(* CODESYS project Syn_Config_2.1.0.library
   Description: Parameter sets the RPP configurator writes and the application takes over (ADR 0017).
   Version: 2.1.0.0
   Title: SynConfig
   Placeholder: SynConfig
   Company: Syntegon Group
   DefaultNamespace: SynConfig

Project tree, tasks and I/O mapping:
  libraries: SynVisu, * (Syntegon Group); Tc2_Standard, * (Beckhoff Automation GmbH)
  DUTs/
    data type E_ConfigAction
    data type E_ConfigCommand
    data type E_ConfigCommandResult
    data type E_ConfigFieldType
    data type E_ConfigResult
    data type ST_ConfigBodyComponent
    data type ST_ConfigBodyComponentParam
    data type ST_ConfigBodyComponentSet
    data type ST_ConfigCartesian
    data type ST_ConfigCartesianParam
    data type ST_ConfigCartesianSet
    data type ST_ConfigCommand
    data type ST_ConfigCommandStatus
    data type ST_ConfigConveyor
    data type ST_ConfigConveyorParam
    data type ST_ConfigConveyorSet
    data type ST_ConfigDelta
    data type ST_ConfigDeltaParam
    data type ST_ConfigDeltaSet
    data type ST_ConfigMachine
    data type ST_ConfigManifest
    data type ST_ConfigManifestEntry
    data type ST_ConfigRecipeField
    data type ST_ConfigRecipeSet
    data type ST_ConfigStaging
    data type ST_ConfigStatus
    data type ST_ConfigXtsGantry
    data type ST_ConfigXtsGantryParam
    data type ST_ConfigXtsGantrySet
    data type ST_ConfigXtsLoop
    data type ST_ConfigXtsLoopParam
    data type ST_ConfigXtsLoopSet
  GVLs/
    global variables CONFIG_GlobalConst
    global variables CONFIG_GlobalConst_Param
  POUs/
    function block _FB_ConfigBodyComponent [ST]: m_Active, m_Cycle, m_PassOnBody, m_Pose
    function block _FB_ConfigCartesian [ST]: m_Active, m_ComponentType, m_Cycle, m_Invalid, m_PassOn, m_Pose
    function block _FB_ConfigComponent [ST]: m_ComponentType, m_Handled, m_Id, m_InvalidFingers, m_InvalidModules, m_InvalidZones, m_PassOnFingers, m_PassOnLimitAreas, m_PassOnModules, m_PassOnZones, m_Register, m_Staging, m_SymbolPath
    function block _FB_ConfigConveyor [ST]: m_Active, m_ComponentType, m_Cycle, m_Invalid, m_PassOn, m_Pose
    function block _FB_ConfigDelta [ST]: m_Active, m_ComponentType, m_Cycle, m_Invalid, m_PassOn, m_Pose, m_Zone, m_ZoneCount
    function block _FB_ConfigMachine [ST]: m_AnswerCommand, m_Command, m_Cycle, m_DeclareField, m_Integer, m_Invalid, m_SetChoice, m_Switch, m_Value
    function block _FB_ConfigSensor [ST]: m_ComponentType, m_PassOn
    function block _FB_ConfigStation [ST]: m_ComponentType, m_PassOn
    function block _FB_ConfigVision [ST]: m_ComponentType, m_PassOn
    function block _FB_ConfigXtsGantry [ST]: m_Active, m_ComponentType, m_Cycle, m_Invalid, m_PassOn, m_Pose
    function block _FB_ConfigXtsLoop [ST]: m_Active, m_ComponentType, m_Cycle, m_Invalid, m_PassOn, m_Pose
    function _FC_GetVersionSynConfig [ST]
*)

// DUTs/E_ConfigAction
{attribute 'qualified_only'}
{attribute 'strict'}
TYPE E_ConfigAction :
(
	(* What a parameter FB does with its staging this cycle (internal). *)
	NONE := 0,
	TAKE_OVER := 1,	// check the staged set and take it over
	RESET := 2		// make the active set invalid: the program values apply again
) UINT;
END_TYPE

// DUTs/E_ConfigCommand
{attribute 'qualified_only'}
{attribute 'strict'}
TYPE E_ConfigCommand :
(
	(* What a machine command asks the application (config protocol 3). Values are part of the gateway contract:
	   append, never renumber. *)
	NONE := 0,
	START := 1,
	STOP := 2,
	RESET := 3
) UINT;
END_TYPE

// DUTs/E_ConfigCommandResult
{attribute 'qualified_only'}
{attribute 'strict'}
TYPE E_ConfigCommandResult :
(
	(* What the application made of the last machine command. Values are part of the gateway contract: append, never
	   renumber. *)
	NONE := 0,		// nothing asked since the PLC started
	ACCEPTED := 1,
	REJECTED := 2	// ST_ConfigCommandStatus.sMessage says why
) UINT;
END_TYPE

// DUTs/E_ConfigFieldType
{attribute 'qualified_only'}
{attribute 'strict'}
TYPE E_ConfigFieldType :
(
	(* How a recipe field's value is kept (config protocol 3). Every value travels as LREAL. Values are part of the
	   gateway contract: append, never renumber. *)
	NUMBER := 0,	// any number within fMin..fMax
	INTEGER := 1,	// a whole number within fMin..fMax, e.g. picks per cycle
	SWITCH := 2,	// on or off: 1 or 0
	CHOICE := 3		// one of the named choices: 0..nChoiceCount-1
) UINT;
END_TYPE

// DUTs/E_ConfigResult
{attribute 'qualified_only'}
{attribute 'strict'}
TYPE E_ConfigResult :
(
	(* What became of the last staged parameter set. Values are part of the gateway contract: append, never renumber. *)
	NONE := 0,		// nothing staged since the PLC started
	PENDING := 1,	// staged, waiting for the application to allow taking it over
	APPLIED := 2,	// taken over (or reset to the program values)
	REJECTED := 3	// not taken over; ST_ConfigStatus.sMessage says why
) UINT;
END_TYPE

// DUTs/ST_ConfigBodyComponent
TYPE ST_ConfigBodyComponent :
STRUCT
	(* vo_Config of _FB_ConfigVision, _FB_ConfigSensor and _FB_ConfigStation: the gateway writes stStaging and
	   stStaged, reads stStatus and stActive. *)
	stStaging : ST_ConfigStaging;
	stStaged : ST_ConfigBodyComponentParam;
	stStatus : ST_ConfigStatus;
	stActive : ST_ConfigBodyComponentParam; // effective values: the active set while one is valid, else the program values
END_STRUCT
END_TYPE

// DUTs/ST_ConfigBodyComponentParam
TYPE ST_ConfigBodyComponentParam :
STRUCT
	(* The parameter set of a component drawn from its bodies (vision system, product sensor, station): what the
	   configurator writes, never its bodies (hardware). Members as in SynVisu.ST_VisuDetectorConfig. *)
	stPose : SynVisu.ST_VisuPose; // MCS
	stOriginShift : SynVisu.ST_VisuPosition; // mm in the component's local frame
	nZoneCount : UINT;
	aZones : ARRAY[0..SynVisu.VISU_GlobalConst_Param.VISU_un_MAX_ZONES - 1] OF SynVisu.ST_VisuZone;
END_STRUCT
END_TYPE

// DUTs/ST_ConfigBodyComponentSet
TYPE ST_ConfigBodyComponentSet :
STRUCT
	(* The active parameter set of a vision system, product sensor or station as the application keeps it, in a
	   VAR PERSISTENT variable passed to m_Cycle of _FB_ConfigVision, _FB_ConfigSensor or _FB_ConfigStation. *)
	bValid : BOOL; // FALSE: no set active, the program values apply
	nVersion : UDINT; // version of stParam
	nLastVersion : UDINT; // last version handed out; versions never repeat, also after a reset
	stParam : ST_ConfigBodyComponentParam;
END_STRUCT
END_TYPE

// DUTs/ST_ConfigCartesian
TYPE ST_ConfigCartesian :
STRUCT
	(* vo_Config of _FB_ConfigCartesian: the gateway writes stStaging and stStaged, reads stStatus and stActive. *)
	stStaging : ST_ConfigStaging;
	stStaged : ST_ConfigCartesianParam;
	stStatus : ST_ConfigStatus;
	stActive : ST_ConfigCartesianParam; // effective values: the active set while one is valid, else the program values
END_STRUCT
END_TYPE

// DUTs/ST_ConfigCartesianParam
TYPE ST_ConfigCartesianParam :
STRUCT
	(* A Cartesian robot's parameter set: what the configurator writes, never its axes, strokes or rail height
	   (hardware). Members as in SynVisu.ST_VisuCartesianConfig. *)
	stPose : SynVisu.ST_VisuPose; // MCS, axis origin X = Y = 0 with Z up
	stOriginShift : SynVisu.ST_VisuPosition; // mm in the robot's local frame
	nZoneCount : UINT;
	aZones : ARRAY[0..SynVisu.VISU_GlobalConst_Param.VISU_un_MAX_ZONES - 1] OF SynVisu.ST_VisuZone;
	nFingerCount : UINT; // gripper fingers with their flange offsets (config protocol 2, ADR 0018)
	aFingers : ARRAY[0..SynVisu.VISU_GlobalConst_Param.VISU_un_MAX_FINGERS - 1] OF SynVisu.ST_VisuFinger;
	stLimitArea : SynVisu.ST_VisuLimitArea; // bActive = FALSE: none
	stTcpLimitArea : SynVisu.ST_VisuLimitArea; // bActive = FALSE: none
END_STRUCT
END_TYPE

// DUTs/ST_ConfigCartesianSet
TYPE ST_ConfigCartesianSet :
STRUCT
	(* A Cartesian robot's active parameter set as the application keeps it, in a VAR PERSISTENT variable passed to
	   _FB_ConfigCartesian.m_Cycle. *)
	bValid : BOOL; // FALSE: no set active, the program values apply
	nVersion : UDINT; // version of stParam
	nLastVersion : UDINT; // last version handed out; versions never repeat, also after a reset
	stParam : ST_ConfigCartesianParam;
END_STRUCT
END_TYPE

// DUTs/ST_ConfigCommand
TYPE ST_ConfigCommand :
STRUCT
	(* A machine command, written by the gateway with bRequested last (config protocol 3). The machine FB clears
	   bRequested once the application answered it. *)
	nCommandId : UDINT; // chosen by the gateway; ST_ConfigCommandStatus.nHandledCommandId names it once answered
	eCommand : E_ConfigCommand;
	bRequested : BOOL; // TRUE: the command waits for the application's answer
END_STRUCT
END_TYPE

// DUTs/ST_ConfigCommandStatus
TYPE ST_ConfigCommandStatus :
STRUCT
	nHandledCommandId : UDINT; // nCommandId of the last command the application answered
	eResult : E_ConfigCommandResult; // what the application made of it
	sMessage : STRING(80); // why it was rejected; empty otherwise
END_STRUCT
END_TYPE

// DUTs/ST_ConfigConveyor
TYPE ST_ConfigConveyor :
STRUCT
	(* vo_Config of _FB_ConfigConveyor: the gateway writes stStaging and stStaged, reads stStatus and stActive. *)
	stStaging : ST_ConfigStaging;
	stStaged : ST_ConfigConveyorParam;
	stStatus : ST_ConfigStatus;
	stActive : ST_ConfigConveyorParam; // effective values: the active set while one is valid, else the program values
END_STRUCT
END_TYPE

// DUTs/ST_ConfigConveyorParam
TYPE ST_ConfigConveyorParam :
STRUCT
	(* A conveyor's parameter set: what the configurator writes, never the belt's length or width (hardware).
	   Members as in SynVisu.ST_VisuConveyorConfig. *)
	stPose : SynVisu.ST_VisuPose; // MCS, belt start on the belt surface; local +X = conveying direction
	stOriginShift : SynVisu.ST_VisuPosition; // mm in the local frame from stPose: origin of the belt coordinates
	nProductTypeCount : UINT;
	aProductTypes : ARRAY[0..SynVisu.VISU_GlobalConst_Param.VISU_un_MAX_PRODUCT_TYPES - 1] OF SynVisu.ST_VisuProductType;
END_STRUCT
END_TYPE

// DUTs/ST_ConfigConveyorSet
TYPE ST_ConfigConveyorSet :
STRUCT
	(* A conveyor's active parameter set as the application keeps it, in a VAR PERSISTENT variable passed to
	   _FB_ConfigConveyor.m_Cycle. *)
	bValid : BOOL; // FALSE: no set active, the program values apply
	nVersion : UDINT; // version of stParam
	nLastVersion : UDINT; // last version handed out; versions never repeat, also after a reset
	stParam : ST_ConfigConveyorParam;
END_STRUCT
END_TYPE

// DUTs/ST_ConfigDelta
TYPE ST_ConfigDelta :
STRUCT
	(* vo_Config of _FB_ConfigDelta: the gateway writes stStaging and stStaged, reads stStatus and stActive. *)
	stStaging : ST_ConfigStaging;
	stStaged : ST_ConfigDeltaParam;
	stStatus : ST_ConfigStatus;
	stActive : ST_ConfigDeltaParam; // effective values: the active set while one is valid, else the program values
END_STRUCT
END_TYPE

// DUTs/ST_ConfigDeltaParam
TYPE ST_ConfigDeltaParam :
STRUCT
	(* A Delta robot's parameter set: what the configurator writes, never its arm geometry (hardware).
	   Members as in SynVisu.ST_VisuDeltaConfig. *)
	stPose : SynVisu.ST_VisuPose; // MCS, base centre
	stOriginShift : SynVisu.ST_VisuPosition; // mm in the base's local frame
	nZoneCount : UINT;
	aZones : ARRAY[0..SynVisu.VISU_GlobalConst_Param.VISU_un_MAX_ZONES - 1] OF SynVisu.ST_VisuZone;
	nFingerCount : UINT; // gripper fingers with their flange offsets (config protocol 2, ADR 0018)
	aFingers : ARRAY[0..SynVisu.VISU_GlobalConst_Param.VISU_un_MAX_FINGERS - 1] OF SynVisu.ST_VisuFinger;
	stWorkingArea : SynVisu.ST_VisuWorkingArea;
	stLimitArea : SynVisu.ST_VisuLimitArea; // bActive = FALSE: none
	stTcpLimitArea : SynVisu.ST_VisuLimitArea; // bActive = FALSE: none
END_STRUCT
END_TYPE

// DUTs/ST_ConfigDeltaSet
TYPE ST_ConfigDeltaSet :
STRUCT
	(* A Delta robot's active parameter set as the application keeps it, in a VAR PERSISTENT variable passed to
	   _FB_ConfigDelta.m_Cycle. *)
	bValid : BOOL; // FALSE: no set active, the program values apply
	nVersion : UDINT; // version of stParam
	nLastVersion : UDINT; // last version handed out; versions never repeat, also after a reset
	stParam : ST_ConfigDeltaParam;
END_STRUCT
END_TYPE

// DUTs/ST_ConfigMachine
TYPE ST_ConfigMachine :
STRUCT
	(* vo_Config of _FB_ConfigMachine (config protocol 3, ADR 0022), listed in the config manifest with id 0 and type
	   NONE. The gateway reads the declared fields once, writes stStaging with aStaged (bStaged or bReset last) and
	   stCommand (bRequested last), and reads stStatus, aActive and stCommandStatus every cycle. Values are kept by
	   field index, every type as LREAL (SWITCH 0 / 1, INTEGER and CHOICE whole numbers). *)
	nFieldCount : UINT; // fields [0..nFieldCount-1] are declared
	aFields : ARRAY[0..CONFIG_GlobalConst_Param.CONFIG_un_MAX_RECIPE_FIELDS - 1] OF ST_ConfigRecipeField;
	stStaging : ST_ConfigStaging;
	aStaged : ARRAY[0..CONFIG_GlobalConst_Param.CONFIG_un_MAX_RECIPE_FIELDS - 1] OF LREAL; // the proposed recipe
	stStatus : ST_ConfigStatus;
	aActive : ARRAY[0..CONFIG_GlobalConst_Param.CONFIG_un_MAX_RECIPE_FIELDS - 1] OF LREAL; // effective values
	stCommand : ST_ConfigCommand;
	stCommandStatus : ST_ConfigCommandStatus;
END_STRUCT
END_TYPE

// DUTs/ST_ConfigManifest
TYPE ST_ConfigManifest :
STRUCT
	(* Where the gateway finds the parameter FBs (ADR 0017). The application declares one instance at the symbol
	   GVL_Config.stManifest; every parameter FB registers itself with m_Register. *)
	nProtocolVersion : UINT := CONFIG_GlobalConst.CONFIG_un_PROTOCOL_VERSION;
	sLibraryVersion : STRING(15); // version of the Syn_Config library actually running, e.g. '1.0.0'
	nCount : UINT; // entries [0..nCount-1] are evaluated
	aEntries : ARRAY[0..CONFIG_GlobalConst_Param.CONFIG_un_MAX_MANIFEST_ENTRIES - 1] OF ST_ConfigManifestEntry;
END_STRUCT
END_TYPE

// DUTs/ST_ConfigManifestEntry
TYPE ST_ConfigManifestEntry :
STRUCT
	nId : UDINT; // manifest id of the Syn_Visu component the parameter FB is for
	eType : SynVisu.E_VisuComponentType; // type of that component
	sPath : STRING(255); // symbol path of the parameter FB's vo_Config, e.g. 'P_Line.fb_InfeedParam.vo_Config'
END_STRUCT
END_TYPE

// DUTs/ST_ConfigRecipeField
TYPE ST_ConfigRecipeField :
STRUCT
	(* One field of the machine's recipe as the application declares it with _FB_ConfigMachine.m_DeclareField
	   (config protocol 3, ADR 0022). The gateway reads the declarations once at discovery. *)
	sName : STRING(31); // unique in the recipe, e.g. 'BeltSpeed'
	nGroup : UDINT; // manifest id of the Syn_Visu component the field belongs to, 0 = the whole machine
	eType : E_ConfigFieldType;
	sUnit : STRING(15); // e.g. 'mm/s', '' = none
	fMin : LREAL; // smallest value of a NUMBER or INTEGER field
	fMax : LREAL; // largest value of a NUMBER or INTEGER field
	fProgramValue : LREAL; // the application's own value, which applies while no recipe is active
	nChoiceCount : UINT; // named values of a CHOICE field
	aChoices : ARRAY[0..CONFIG_GlobalConst_Param.CONFIG_un_MAX_CHOICES - 1] OF STRING(31); // their names, from value 0
END_STRUCT
END_TYPE

// DUTs/ST_ConfigRecipeSet
TYPE ST_ConfigRecipeSet :
STRUCT
	(* The machine's active recipe as the application keeps it, in a VAR PERSISTENT variable passed to
	   _FB_ConfigMachine.m_Cycle. Values by field index: keep the fields' order, add new ones at the end. *)
	bValid : BOOL; // FALSE: no recipe active, the program values apply
	nVersion : UDINT; // version of aValues
	nLastVersion : UDINT; // last version handed out; versions never repeat, also after a reset
	aValues : ARRAY[0..CONFIG_GlobalConst_Param.CONFIG_un_MAX_RECIPE_FIELDS - 1] OF LREAL;
END_STRUCT
END_TYPE

// DUTs/ST_ConfigStaging
TYPE ST_ConfigStaging :
STRUCT
	(* Written by the gateway in one ADS sum-write, bStaged or bReset last, so a set is never seen staged half
	   written (ADR 0017). The parameter FB clears bStaged and bReset once it handled them. *)
	nBaseVersion : UDINT; // active version the staged set is based on; another active version rejects it
	nStageId : UDINT; // chosen by the gateway; ST_ConfigStatus.nHandledStageId names it once handled
	bReset : BOOL; // TRUE: make the active set invalid, the program values apply again
	bStaged : BOOL; // TRUE: stStaged is complete and waits to be taken over
END_STRUCT
END_TYPE

// DUTs/ST_ConfigStatus
TYPE ST_ConfigStatus :
STRUCT
	nActiveVersion : UDINT; // version of the active set; 0 while the program values apply
	nHandledStageId : UDINT; // nStageId of the last staging handled (taken over, rejected or reset)
	eResult : E_ConfigResult; // what became of it
	sMessage : STRING(80); // why it was rejected; empty otherwise
END_STRUCT
END_TYPE

// DUTs/ST_ConfigXtsGantry
TYPE ST_ConfigXtsGantry :
STRUCT
	(* vo_Config of _FB_ConfigXtsGantry: the gateway writes stStaging and stStaged, reads stStatus and stActive. *)
	stStaging : ST_ConfigStaging;
	stStaged : ST_ConfigXtsGantryParam;
	stStatus : ST_ConfigStatus;
	stActive : ST_ConfigXtsGantryParam; // effective values: the active set while one is valid, else the program values
END_STRUCT
END_TYPE

// DUTs/ST_ConfigXtsGantryParam
TYPE ST_ConfigXtsGantryParam :
STRUCT
	(* An XTS gantry's parameter set: what the configurator writes, never its strokes, tool offsets or mover size
	   (hardware). Members as in SynVisu.ST_VisuXtsGantryConfig. *)
	stPose : SynVisu.ST_VisuPose; // MCS, track start on top of the movers with Z = 0
	stOriginShift : SynVisu.ST_VisuPosition; // mm in the track's local frame
	nModuleCount : UINT;
	aModules : ARRAY[0..SynVisu.VISU_GlobalConst_Param.VISU_un_MAX_MODULES - 1] OF SynVisu.ST_VisuTrackModule;
	nZoneCount : UINT;
	aZones : ARRAY[0..SynVisu.VISU_GlobalConst_Param.VISU_un_MAX_ZONES - 1] OF SynVisu.ST_VisuZone;
	nFingerCount : UINT; // gripper fingers of every mover, with their flange offsets (config protocol 2, ADR 0018)
	aFingers : ARRAY[0..SynVisu.VISU_GlobalConst_Param.VISU_un_MAX_FINGERS - 1] OF SynVisu.ST_VisuFinger;
	stLimitArea : SynVisu.ST_VisuLimitArea; // bActive = FALSE: none
	stTcpLimitArea : SynVisu.ST_VisuLimitArea; // bActive = FALSE: none
END_STRUCT
END_TYPE

// DUTs/ST_ConfigXtsGantrySet
TYPE ST_ConfigXtsGantrySet :
STRUCT
	(* An XTS gantry's active parameter set as the application keeps it, in a VAR PERSISTENT variable passed to
	   _FB_ConfigXtsGantry.m_Cycle. *)
	bValid : BOOL; // FALSE: no set active, the program values apply
	nVersion : UDINT; // version of stParam
	nLastVersion : UDINT; // last version handed out; versions never repeat, also after a reset
	stParam : ST_ConfigXtsGantryParam;
END_STRUCT
END_TYPE

// DUTs/ST_ConfigXtsLoop
TYPE ST_ConfigXtsLoop :
STRUCT
	(* vo_Config of _FB_ConfigXtsLoop: the gateway writes stStaging and stStaged, reads stStatus and stActive. *)
	stStaging : ST_ConfigStaging;
	stStaged : ST_ConfigXtsLoopParam;
	stStatus : ST_ConfigStatus;
	stActive : ST_ConfigXtsLoopParam; // effective values: the active set while one is valid, else the program values
END_STRUCT
END_TYPE

// DUTs/ST_ConfigXtsLoopParam
TYPE ST_ConfigXtsLoopParam :
STRUCT
	(* An XTS loop's parameter set: what the configurator writes, never its tool offset or mover size (hardware).
	   Members as in SynVisu.ST_VisuXtsLoopConfig. *)
	stPose : SynVisu.ST_VisuPose; // MCS, start of module 1
	stOriginShift : SynVisu.ST_VisuPosition; // mm in the loop's local frame
	nModuleCount : UINT;
	aModules : ARRAY[0..SynVisu.VISU_GlobalConst_Param.VISU_un_MAX_MODULES - 1] OF SynVisu.ST_VisuTrackModule;
	nZoneCount : UINT;
	aZones : ARRAY[0..SynVisu.VISU_GlobalConst_Param.VISU_un_MAX_ZONES - 1] OF SynVisu.ST_VisuZone;
	nFingerCount : UINT; // gripper fingers of every mover, with their flange offsets (config protocol 2, ADR 0018)
	aFingers : ARRAY[0..SynVisu.VISU_GlobalConst_Param.VISU_un_MAX_FINGERS - 1] OF SynVisu.ST_VisuFinger;
END_STRUCT
END_TYPE

// DUTs/ST_ConfigXtsLoopSet
TYPE ST_ConfigXtsLoopSet :
STRUCT
	(* An XTS loop's active parameter set as the application keeps it, in a VAR PERSISTENT variable passed to
	   _FB_ConfigXtsLoop.m_Cycle. *)
	bValid : BOOL; // FALSE: no set active, the program values apply
	nVersion : UDINT; // version of stParam
	nLastVersion : UDINT; // last version handed out; versions never repeat, also after a reset
	stParam : ST_ConfigXtsLoopParam;
END_STRUCT
END_TYPE

// GVLs/CONFIG_GlobalConst
(****************************************************************************************************<br>
© Syntegon Group.<br>
All rights reserved, also regarding any disposal, exploitation, reproduction, editing, distribution,<br>
as well as in the event of applications for industrial property rights.<br>
*****************************************************************************************************<br>
DESCRIPTION:<br>
Global constants of the Syn_Config library.<br>
****************************************************************************************************)
{attribute 'qualified_only'}
VAR_GLOBAL CONSTANT
	(* Version of the Syn_Config <-> gateway contract (ADR 0017). The gateway writes nothing to a PLC whose config
	   manifest reports a version it does not know (it knows 2 and 3). Bump together with CONFIG_PROTOCOL_VERSION in
	   the gateway.
	   1: conveyor (pose, origin shift, product types) and Delta (pose, origin shift, zones, working, limit and
	      TCP limit area); since library 1.1.0 also XTS gantry, XTS loop, Cartesian, vision, sensor and station
	      (new parameter FBs only: no change for a gateway or an application of 1.0.0).
	   2: gripper fingers with their flange offsets (nFingerCount, aFingers) in the parameter sets of the Delta,
	      the XTS gantry and loop and the Cartesian robot (library 2.0.0, ADR 0018).
	   3: the machine FB _FB_ConfigMachine (id 0, type NONE in the manifest): recipe fields the application declares,
	      their staging, and machine commands (library 2.1.0, ADR 0022). A PLC of version 2 still gets its parameter
	      sets written, but no recipe and no commands. *)
	CONFIG_un_PROTOCOL_VERSION			: UINT := 3;
	(* Version of this library (config manifest sLibraryVersion). Bump together with _FC_GetVersionSynConfig and the
	   project version. *)
	CONFIG_str_LIBRARY_VERSION			: STRING(15) := '2.1.0';
END_VAR

// GVLs/CONFIG_GlobalConst_Param
(****************************************************************************************************<br>
© Syntegon Group.<br>
All rights reserved, also regarding any disposal, exploitation, reproduction, editing, distribution,<br>
as well as in the event of applications for industrial property rights.<br>
*****************************************************************************************************<br>
DESCRIPTION:<br>
Library parameters of Syn_Config: array sizes of the interface structures. The lists of a parameter set have the
sizes of Syn_Visu's (VISU_GlobalConst_Param), so every set fits the visualisation it is passed on to.<br>
****************************************************************************************************)
{attribute 'qualified_only'}
VAR_GLOBAL CONSTANT
	CONFIG_un_MAX_MANIFEST_ENTRIES		: UINT := 32;	// [-] parameter FBs in the config manifest
	CONFIG_un_MAX_RECIPE_FIELDS			: UINT := 64;	// [-] fields of the machine's recipe (_FB_ConfigMachine)
	CONFIG_un_MAX_CHOICES				: UINT := 8;	// [-] named values of a CHOICE recipe field
END_VAR

// POUs/_FB_ConfigBodyComponent
(****************************************************************************************************<br>
© Syntegon Group.<br>
All rights reserved, also regarding any disposal, exploitation, reproduction, editing, distribution,<br>
as well as in the event of applications for industrial property rights.<br>
*****************************************************************************************************<br>
DESCRIPTION:<br>
Base of the parameter FBs of components drawn from their bodies (_FB_ConfigVision, _FB_ConfigSensor,<br>
_FB_ConfigStation, ADR 0017): their pose, origin shift and zones, written by the configurator, taken over when<br>
the application allows it. The bodies are hardware and stay the application's. Typical cycle:<br>
  fb_VisionParam.m_Register(vio_Manifest := GVL_Config.stManifest, vi_udn_Id := fb_Vision.m_Id());<br>
  fb_VisionParam.m_Cycle(vio_Default := VisionDefault, vio_Set := VisionSet, vi_b_ApplyAllowed := b_Stopped);<br>
  fb_Vision.m_Configure(vi_Pose := fb_VisionParam.m_Pose(), vi_lr_FieldLength := 400, ...);<br>
  fb_VisionParam.m_PassOn(vio_Visu := fb_Vision);<br>
Not used directly.<br>
*****************************************************************************************************<br>
OUTPUT VALUES:<br>
vo_Config is the contract structure the gateway reads and writes at the path in the config manifest.<br>
*****************************************************************************************************<br>
VERSION         ¦ DATE       ¦ NAME      ¦ CHANGE<br>
Syn_Config 1.1.0 ¦ 2026-11-10 ¦ J.Willner ¦ New<br>
****************************************************************************************************)
FUNCTION_BLOCK ABSTRACT _FB_ConfigBodyComponent EXTENDS _FB_ConfigComponent
VAR_OUTPUT
	vo_Config							: ST_ConfigBodyComponent;	// contract structure of the gateway
END_VAR

(****************************************************************************************************<br>
© Syntegon Group.<br>
All rights reserved, also regarding any disposal, exploitation, reproduction, editing, distribution,<br>
as well as in the event of applications for industrial property rights.<br>
*****************************************************************************************************<br>
DESCRIPTION:<br>
All effective values (zones, ...), for the application's own logic.<br>
****************************************************************************************************)
METHOD m_Active : ST_ConfigBodyComponentParam
m_Active := vo_Config.stActive;
END_METHOD

(****************************************************************************************************<br>
© Syntegon Group.<br>
All rights reserved, also regarding any disposal, exploitation, reproduction, editing, distribution,<br>
as well as in the event of applications for industrial property rights.<br>
*****************************************************************************************************<br>
DESCRIPTION:<br>
Every cycle: handles a staged set or a reset (a set only while vi_b_ApplyAllowed), keeps the active set in<br>
vio_Set and gives the effective values in vo_Config.stActive: the active set while one is valid, else the<br>
program values vio_Default.<br>
*****************************************************************************************************<br>
OUTPUT VALUES:<br>
TRUE in the cycle a set was taken over or reset.<br>
****************************************************************************************************)
METHOD m_Cycle : BOOL
VAR_IN_OUT CONSTANT
	vio_Default							: ST_ConfigBodyComponentParam;	// the application's program values
END_VAR
VAR_IN_OUT
	vio_Set								: ST_ConfigBodyComponentSet;	// the application's VAR PERSISTENT active set
END_VAR
VAR_INPUT
	vi_b_ApplyAllowed					: BOOL;	// [-] a staged set may be taken over now, e.g. while the machine stands
END_VAR
VAR
	str_TempRejection					: STRING(80);
END_VAR
m_Cycle := FALSE;
CASE m_Staging(vio_Staging := vo_Config.stStaging, vio_Status := vo_Config.stStatus, vi_b_ApplyAllowed := vi_b_ApplyAllowed,
	vi_udn_ActiveVersion := SEL(vio_Set.bValid, 0, vio_Set.nVersion)) OF
	E_ConfigAction.RESET:
		vio_Set.bValid := FALSE;
		m_Handled(vio_Staging := vo_Config.stStaging, vio_Status := vo_Config.stStatus, vi_str_Rejection := '');
		m_Cycle := TRUE;
	E_ConfigAction.TAKE_OVER:
		str_TempRejection := m_InvalidZones(vio_aZones := vo_Config.stStaged.aZones, vi_un_Count := vo_Config.stStaged.nZoneCount);
		IF str_TempRejection = '' THEN
			vio_Set.nLastVersion := vio_Set.nLastVersion + 1;
			vio_Set.nVersion := vio_Set.nLastVersion;
			vio_Set.stParam := vo_Config.stStaged;
			vio_Set.bValid := TRUE;
			m_Cycle := TRUE;
		END_IF
		m_Handled(vio_Staging := vo_Config.stStaging, vio_Status := vo_Config.stStatus, vi_str_Rejection := str_TempRejection);
END_CASE


(****************************************************************************************************
EFFECTIVE VALUES
****************************************************************************************************)
IF vio_Set.bValid THEN
	vo_Config.stActive := vio_Set.stParam;
	vo_Config.stStatus.nActiveVersion := vio_Set.nVersion;
ELSE
	vo_Config.stActive := vio_Default;
	vo_Config.stStatus.nActiveVersion := 0;
END_IF
END_METHOD

(****************************************************************************************************<br>
© Syntegon Group.<br>
All rights reserved, also regarding any disposal, exploitation, reproduction, editing, distribution,<br>
as well as in the event of applications for industrial property rights.<br>
*****************************************************************************************************<br>
DESCRIPTION:<br>
Passes the effective origin shift and zones on to the component's Syn_Visu FB; for m_PassOn of the derived FB,<br>
which knows where the visualisation keeps its zone count.<br>
****************************************************************************************************)
METHOD PROTECTED m_PassOnBody : BOOL
VAR_IN_OUT
	vio_Visu							: SynVisu._FB_VisuBodyComponent;	// the component's Syn_Visu FB
END_VAR
VAR_INPUT
	vi_un_VisuZoneCount					: UINT;	// [-] zones the visualisation has now, its stConfig.nZoneCount
END_VAR
m_PassOnBody := TRUE;
vio_Visu.m_SetOriginShift(vi_lr_X := vo_Config.stActive.stOriginShift.fX, vi_lr_Y := vo_Config.stActive.stOriginShift.fY,
	vi_lr_Z := vo_Config.stActive.stOriginShift.fZ);
m_PassOnZones(vio_Visu := vio_Visu, vio_aZones := vo_Config.stActive.aZones, vi_un_Count := vo_Config.stActive.nZoneCount,
	vi_un_VisuCount := vi_un_VisuZoneCount);
END_METHOD

(****************************************************************************************************<br>
© Syntegon Group.<br>
All rights reserved, also regarding any disposal, exploitation, reproduction, editing, distribution,<br>
as well as in the event of applications for industrial property rights.<br>
*****************************************************************************************************<br>
DESCRIPTION:<br>
Effective pose (MCS), for the application's logic and its Syn_Visu m_Configure call.<br>
****************************************************************************************************)
METHOD m_Pose : SynVisu.ST_VisuPose
m_Pose := vo_Config.stActive.stPose;
END_METHOD

END_FUNCTION_BLOCK

// POUs/_FB_ConfigVision
(****************************************************************************************************<br>
© Syntegon Group.<br>
All rights reserved, also regarding any disposal, exploitation, reproduction, editing, distribution,<br>
as well as in the event of applications for industrial property rights.<br>
*****************************************************************************************************<br>
DESCRIPTION:<br>
Parameter set of one vision system (ADR 0017): its pose, origin shift and zones. See _FB_ConfigBodyComponent.<br>
*****************************************************************************************************<br>
VERSION         ¦ DATE       ¦ NAME      ¦ CHANGE<br>
Syn_Config 1.1.0 ¦ 2026-11-10 ¦ J.Willner ¦ New<br>
****************************************************************************************************)
FUNCTION_BLOCK _FB_ConfigVision EXTENDS _FB_ConfigBodyComponent

(****************************************************************************************************<br>
© Syntegon Group.<br>
All rights reserved, also regarding any disposal, exploitation, reproduction, editing, distribution,<br>
as well as in the event of applications for industrial property rights.<br>
*****************************************************************************************************<br>
DESCRIPTION:<br>
A vision system.<br>
****************************************************************************************************)
METHOD PROTECTED m_ComponentType : SynVisu.E_VisuComponentType
m_ComponentType := SynVisu.E_VisuComponentType.VISION;
END_METHOD

(****************************************************************************************************<br>
© Syntegon Group.<br>
All rights reserved, also regarding any disposal, exploitation, reproduction, editing, distribution,<br>
as well as in the event of applications for industrial property rights.<br>
*****************************************************************************************************<br>
DESCRIPTION:<br>
Passes the effective origin shift and zones on to the vision system's Syn_Visu FB. The pose goes with the<br>
application's own m_Configure call (with the field of view, hardware): vi_Pose := m_Pose(). Call it after<br>
m_Cycle, every cycle.<br>
****************************************************************************************************)
METHOD m_PassOn : BOOL
VAR_IN_OUT
	vio_Visu							: SynVisu._FB_VisuVision;	// the vision system's Syn_Visu FB
END_VAR
m_PassOn := m_PassOnBody(vio_Visu := vio_Visu, vi_un_VisuZoneCount := vio_Visu.vo_Visu.stConfig.nZoneCount);
END_METHOD

END_FUNCTION_BLOCK

// POUs/_FB_ConfigSensor
(****************************************************************************************************<br>
© Syntegon Group.<br>
All rights reserved, also regarding any disposal, exploitation, reproduction, editing, distribution,<br>
as well as in the event of applications for industrial property rights.<br>
*****************************************************************************************************<br>
DESCRIPTION:<br>
Parameter set of one product sensor (ADR 0017): its pose, origin shift and zones. See _FB_ConfigBodyComponent.<br>
*****************************************************************************************************<br>
VERSION         ¦ DATE       ¦ NAME      ¦ CHANGE<br>
Syn_Config 1.1.0 ¦ 2026-11-10 ¦ J.Willner ¦ New<br>
****************************************************************************************************)
FUNCTION_BLOCK _FB_ConfigSensor EXTENDS _FB_ConfigBodyComponent

(****************************************************************************************************<br>
© Syntegon Group.<br>
All rights reserved, also regarding any disposal, exploitation, reproduction, editing, distribution,<br>
as well as in the event of applications for industrial property rights.<br>
*****************************************************************************************************<br>
DESCRIPTION:<br>
A product sensor.<br>
****************************************************************************************************)
METHOD PROTECTED m_ComponentType : SynVisu.E_VisuComponentType
m_ComponentType := SynVisu.E_VisuComponentType.SENSOR;
END_METHOD

(****************************************************************************************************<br>
© Syntegon Group.<br>
All rights reserved, also regarding any disposal, exploitation, reproduction, editing, distribution,<br>
as well as in the event of applications for industrial property rights.<br>
*****************************************************************************************************<br>
DESCRIPTION:<br>
Passes the effective origin shift and zones on to the sensor's Syn_Visu FB. The pose goes with the<br>
application's own m_Configure call (with the beam length, hardware): vi_Pose := m_Pose(). Call it after<br>
m_Cycle, every cycle.<br>
****************************************************************************************************)
METHOD m_PassOn : BOOL
VAR_IN_OUT
	vio_Visu							: SynVisu._FB_VisuSensor;	// the sensor's Syn_Visu FB
END_VAR
m_PassOn := m_PassOnBody(vio_Visu := vio_Visu, vi_un_VisuZoneCount := vio_Visu.vo_Visu.stConfig.nZoneCount);
END_METHOD

END_FUNCTION_BLOCK

// POUs/_FB_ConfigStation
(****************************************************************************************************<br>
© Syntegon Group.<br>
All rights reserved, also regarding any disposal, exploitation, reproduction, editing, distribution,<br>
as well as in the event of applications for industrial property rights.<br>
*****************************************************************************************************<br>
DESCRIPTION:<br>
Parameter set of one station (reject unit, labeller, ..., ADR 0017): its pose, origin shift and zones. See<br>
_FB_ConfigBodyComponent.<br>
*****************************************************************************************************<br>
VERSION         ¦ DATE       ¦ NAME      ¦ CHANGE<br>
Syn_Config 1.1.0 ¦ 2026-11-10 ¦ J.Willner ¦ New<br>
****************************************************************************************************)
FUNCTION_BLOCK _FB_ConfigStation EXTENDS _FB_ConfigBodyComponent

(****************************************************************************************************<br>
© Syntegon Group.<br>
All rights reserved, also regarding any disposal, exploitation, reproduction, editing, distribution,<br>
as well as in the event of applications for industrial property rights.<br>
*****************************************************************************************************<br>
DESCRIPTION:<br>
A station.<br>
****************************************************************************************************)
METHOD PROTECTED m_ComponentType : SynVisu.E_VisuComponentType
m_ComponentType := SynVisu.E_VisuComponentType.STATION;
END_METHOD

(****************************************************************************************************<br>
© Syntegon Group.<br>
All rights reserved, also regarding any disposal, exploitation, reproduction, editing, distribution,<br>
as well as in the event of applications for industrial property rights.<br>
*****************************************************************************************************<br>
DESCRIPTION:<br>
Passes the effective origin shift and zones on to the station's Syn_Visu FB. The pose goes with the<br>
application's own m_Configure call: vi_Pose := m_Pose(); its bodies stay the application's (hardware). Call it<br>
after m_Cycle, every cycle.<br>
****************************************************************************************************)
METHOD m_PassOn : BOOL
VAR_IN_OUT
	vio_Visu							: SynVisu._FB_VisuStation;	// the station's Syn_Visu FB
END_VAR
m_PassOn := m_PassOnBody(vio_Visu := vio_Visu, vi_un_VisuZoneCount := vio_Visu.vo_Visu.stConfig.nZoneCount);
END_METHOD

END_FUNCTION_BLOCK

// POUs/_FB_ConfigComponent
(****************************************************************************************************<br>
© Syntegon Group.<br>
All rights reserved, also regarding any disposal, exploitation, reproduction, editing, distribution,<br>
as well as in the event of applications for industrial property rights.<br>
*****************************************************************************************************<br>
DESCRIPTION:<br>
Base of every parameter FB (_FB_ConfigConveyor, _FB_ConfigDelta, _FB_ConfigXtsGantry, ...): the config<br>
manifest entry, what is done with a staging (ADR 0017) and the helpers for zones, fingers, limit areas and<br>
track modules the derived FBs share. Not used directly.<br>
*****************************************************************************************************<br>
VERSION         ¦ DATE       ¦ NAME      ¦ CHANGE<br>
Syn_Config 1.0.0 ¦ 2026-11-10 ¦ J.Willner ¦ First version: conveyor and Delta<br>
Syn_Config 1.1.0 ¦ 2026-11-10 ¦ J.Willner ¦ Helpers m_PassOn..., m_Invalid... for every type<br>
Syn_Config 2.0.0 ¦ 2026-11-11 ¦ J.Willner ¦ m_InvalidFingers, m_PassOnFingers (ADR 0018)<br>
****************************************************************************************************)
{attribute 'reflection'}
FUNCTION_BLOCK ABSTRACT _FB_ConfigComponent
VAR
	udn_ComponentId						: UDINT;	// [-] id of the Syn_Visu component, 0 = not registered
	(* Device tree path of this instance, e.g. 'RPP_Visu.Syn_Visu_Demo.P_VisuDemoDelta.fb_InfeedParam', set by TwinCAT
	   at initialisation. *)
	{attribute 'instance-path'}
	{attribute 'noinit'}
	str_InstancePath					: STRING(255);
	str_SymbolPath						: STRING(255);	// symbol path of vo_Config for the manifest, from str_InstancePath
END_VAR

(****************************************************************************************************<br>
© Syntegon Group.<br>
All rights reserved, also regarding any disposal, exploitation, reproduction, editing, distribution,<br>
as well as in the event of applications for industrial property rights.<br>
*****************************************************************************************************<br>
DESCRIPTION:<br>
Type of the Syn_Visu component this FB parametrises. Overridden by every derived FB.<br>
****************************************************************************************************)
METHOD PROTECTED m_ComponentType : SynVisu.E_VisuComponentType
m_ComponentType := SynVisu.E_VisuComponentType.NONE;
END_METHOD

(****************************************************************************************************<br>
© Syntegon Group.<br>
All rights reserved, also regarding any disposal, exploitation, reproduction, editing, distribution,<br>
as well as in the event of applications for industrial property rights.<br>
*****************************************************************************************************<br>
DESCRIPTION:<br>
Reports the staging as handled: taken over (or reset) with an empty vi_str_Rejection, else rejected for that<br>
reason. Clears bStaged and bReset. TRUE when taken over.<br>
****************************************************************************************************)
METHOD PROTECTED m_Handled : BOOL
VAR_IN_OUT
	vio_Staging							: ST_ConfigStaging;	// vo_Config.stStaging
	vio_Status							: ST_ConfigStatus;	// vo_Config.stStatus
END_VAR
VAR_INPUT
	vi_str_Rejection					: STRING(80);	// why the set is not taken over; '' = taken over
END_VAR
m_Handled := vi_str_Rejection = '';
vio_Status.nHandledStageId := vio_Staging.nStageId;
IF m_Handled THEN
	vio_Status.eResult := E_ConfigResult.APPLIED;
	vio_Status.sMessage := '';
ELSE
	vio_Status.eResult := E_ConfigResult.REJECTED;
	vio_Status.sMessage := vi_str_Rejection;
END_IF
vio_Staging.bStaged := FALSE;
vio_Staging.bReset := FALSE;
END_METHOD

(****************************************************************************************************<br>
© Syntegon Group.<br>
All rights reserved, also regarding any disposal, exploitation, reproduction, editing, distribution,<br>
as well as in the event of applications for industrial property rights.<br>
*****************************************************************************************************<br>
DESCRIPTION:<br>
Id given to m_Register (the Syn_Visu component's id); 0 while not registered.<br>
****************************************************************************************************)
METHOD m_Id : UDINT
m_Id := udn_ComponentId;
END_METHOD

(****************************************************************************************************<br>
© Syntegon Group.<br>
All rights reserved, also regarding any disposal, exploitation, reproduction, editing, distribution,<br>
as well as in the event of applications for industrial property rights.<br>
*****************************************************************************************************<br>
DESCRIPTION:<br>
Why a staged set's gripper fingers cannot be taken over; '' when they can: more fingers than the list holds, or<br>
a finger without a diameter or height.<br>
****************************************************************************************************)
METHOD PROTECTED m_InvalidFingers : STRING(80)
VAR_IN_OUT CONSTANT
	(* staged fingers *)
	vio_aFingers						: ARRAY[0..SynVisu.VISU_GlobalConst_Param.VISU_un_MAX_FINGERS - 1] OF SynVisu.ST_VisuFinger;
END_VAR
VAR_INPUT
	vi_un_Count							: UINT;	// [-] staged fingers in vio_aFingers
END_VAR
VAR
	un_TempIndex						: UINT;
END_VAR
m_InvalidFingers := '';
IF vi_un_Count > SynVisu.VISU_GlobalConst_Param.VISU_un_MAX_FINGERS THEN
	m_InvalidFingers := CONCAT('More than ', CONCAT(UINT_TO_STRING(SynVisu.VISU_GlobalConst_Param.VISU_un_MAX_FINGERS), ' fingers'));
	RETURN;
END_IF
un_TempIndex := 0;
WHILE un_TempIndex < vi_un_Count DO
	IF vio_aFingers[un_TempIndex].fDiameter <= 0 OR vio_aFingers[un_TempIndex].fHeight <= 0 THEN
		m_InvalidFingers := CONCAT('Finger ', CONCAT(UINT_TO_STRING(un_TempIndex + 1), ' has no diameter or height'));
		RETURN;
	END_IF
	un_TempIndex := un_TempIndex + 1;
END_WHILE
END_METHOD

(****************************************************************************************************<br>
© Syntegon Group.<br>
All rights reserved, also regarding any disposal, exploitation, reproduction, editing, distribution,<br>
as well as in the event of applications for industrial property rights.<br>
*****************************************************************************************************<br>
DESCRIPTION:<br>
Why a staged set's track modules cannot be taken over; '' when they can: more modules than the list holds,<br>
none at all, or a module without a length.<br>
****************************************************************************************************)
METHOD PROTECTED m_InvalidModules : STRING(80)
VAR_IN_OUT CONSTANT
	(* staged modules *)
	vio_aModules						: ARRAY[0..SynVisu.VISU_GlobalConst_Param.VISU_un_MAX_MODULES - 1] OF SynVisu.ST_VisuTrackModule;
END_VAR
VAR_INPUT
	vi_un_Count							: UINT;	// [-] staged modules in vio_aModules
END_VAR
VAR
	un_TempIndex						: UINT;
END_VAR
m_InvalidModules := '';
IF vi_un_Count > SynVisu.VISU_GlobalConst_Param.VISU_un_MAX_MODULES THEN
	m_InvalidModules := CONCAT('More than ', CONCAT(UINT_TO_STRING(SynVisu.VISU_GlobalConst_Param.VISU_un_MAX_MODULES), ' track modules'));
	RETURN;
END_IF
IF vi_un_Count = 0 THEN
	m_InvalidModules := 'A track without modules';
	RETURN;
END_IF
un_TempIndex := 0;
WHILE un_TempIndex < vi_un_Count DO
	IF vio_aModules[un_TempIndex].fLength <= 0 THEN
		m_InvalidModules := CONCAT('Track module ', CONCAT(UINT_TO_STRING(un_TempIndex + 1), ' has no length'));
		RETURN;
	END_IF
	un_TempIndex := un_TempIndex + 1;
END_WHILE
END_METHOD

(****************************************************************************************************<br>
© Syntegon Group.<br>
All rights reserved, also regarding any disposal, exploitation, reproduction, editing, distribution,<br>
as well as in the event of applications for industrial property rights.<br>
*****************************************************************************************************<br>
DESCRIPTION:<br>
Why a staged set's zones cannot be taken over; '' when they can: more zones than the list holds, or a zone on<br>
no conveyor (id 0).<br>
****************************************************************************************************)
METHOD PROTECTED m_InvalidZones : STRING(80)
VAR_IN_OUT CONSTANT
	(* staged zones *)
	vio_aZones							: ARRAY[0..SynVisu.VISU_GlobalConst_Param.VISU_un_MAX_ZONES - 1] OF SynVisu.ST_VisuZone;
END_VAR
VAR_INPUT
	vi_un_Count							: UINT;	// [-] staged zones in vio_aZones
END_VAR
VAR
	un_TempIndex						: UINT;
END_VAR
m_InvalidZones := '';
IF vi_un_Count > SynVisu.VISU_GlobalConst_Param.VISU_un_MAX_ZONES THEN
	m_InvalidZones := CONCAT('More than ', CONCAT(UINT_TO_STRING(SynVisu.VISU_GlobalConst_Param.VISU_un_MAX_ZONES), ' zones'));
	RETURN;
END_IF
un_TempIndex := 0;
WHILE un_TempIndex < vi_un_Count DO
	IF vio_aZones[un_TempIndex].nConveyorId = 0 THEN
		m_InvalidZones := CONCAT('Zone ', CONCAT(UINT_TO_STRING(un_TempIndex + 1), ' lies on no conveyor'));
		RETURN;
	END_IF
	un_TempIndex := un_TempIndex + 1;
END_WHILE
END_METHOD

(****************************************************************************************************<br>
© Syntegon Group.<br>
All rights reserved, also regarding any disposal, exploitation, reproduction, editing, distribution,<br>
as well as in the event of applications for industrial property rights.<br>
*****************************************************************************************************<br>
DESCRIPTION:<br>
Passes the effective gripper fingers with their flange offsets on to a robot's Syn_Visu FB (ADR 0018). Syn_Visu's<br>
finger count only grows: the fingers are cleared first only when the set has fewer than the visualisation, so<br>
its config version only changes when a value does.<br>
****************************************************************************************************)
METHOD PROTECTED m_PassOnFingers : BOOL
VAR_IN_OUT
	vio_Visu							: SynVisu._FB_VisuRobot;	// the robot's Syn_Visu FB
END_VAR
VAR_IN_OUT CONSTANT
	(* effective fingers *)
	vio_aFingers						: ARRAY[0..SynVisu.VISU_GlobalConst_Param.VISU_un_MAX_FINGERS - 1] OF SynVisu.ST_VisuFinger;
END_VAR
VAR_INPUT
	vi_un_Count							: UINT;	// [-] effective fingers in vio_aFingers
	vi_un_VisuCount						: UINT;	// [-] fingers the visualisation has now, its stConfig.nFingerCount
END_VAR
VAR
	un_TempIndex						: UINT;
END_VAR
m_PassOnFingers := TRUE;
IF vi_un_VisuCount > vi_un_Count THEN
	vio_Visu.m_ClearFingers();
END_IF
un_TempIndex := 0;
WHILE un_TempIndex < vi_un_Count AND un_TempIndex < SynVisu.VISU_GlobalConst_Param.VISU_un_MAX_FINGERS DO
	vio_Visu.m_SetFinger(vi_un_Finger := un_TempIndex + 1, vi_lr_Diameter := vio_aFingers[un_TempIndex].fDiameter,
		vi_lr_Height := vio_aFingers[un_TempIndex].fHeight);
	vio_Visu.m_SetFingerOffset(vi_un_Finger := un_TempIndex + 1, vi_lr_X := vio_aFingers[un_TempIndex].stOffset.fX,
		vi_lr_Y := vio_aFingers[un_TempIndex].stOffset.fY, vi_lr_Z := vio_aFingers[un_TempIndex].stOffset.fZ,
		vi_lr_Rz := vio_aFingers[un_TempIndex].stOffset.fRz);
	un_TempIndex := un_TempIndex + 1;
END_WHILE
END_METHOD

(****************************************************************************************************<br>
© Syntegon Group.<br>
All rights reserved, also regarding any disposal, exploitation, reproduction, editing, distribution,<br>
as well as in the event of applications for industrial property rights.<br>
*****************************************************************************************************<br>
DESCRIPTION:<br>
Passes the effective limit area and TCP limit area on to a robot's Syn_Visu FB (Delta, XTS gantry, Cartesian);<br>
an area with bActive = FALSE is cleared.<br>
****************************************************************************************************)
METHOD PROTECTED m_PassOnLimitAreas : BOOL
VAR_IN_OUT
	vio_Visu							: SynVisu._FB_VisuRobot;	// the robot's Syn_Visu FB
END_VAR
VAR_IN_OUT CONSTANT
	vio_LimitArea						: SynVisu.ST_VisuLimitArea;	// effective limit area
	vio_TcpLimitArea					: SynVisu.ST_VisuLimitArea;	// effective TCP limit area
END_VAR
m_PassOnLimitAreas := TRUE;
IF vio_LimitArea.bActive THEN
	vio_Visu.m_SetLimitArea(vi_lr_XMin := vio_LimitArea.fXMin, vi_lr_XMax := vio_LimitArea.fXMax,
		vi_lr_YMin := vio_LimitArea.fYMin, vi_lr_YMax := vio_LimitArea.fYMax,
		vi_lr_ZMin := vio_LimitArea.fZMin, vi_lr_ZMax := vio_LimitArea.fZMax);
ELSE
	vio_Visu.m_ClearLimitArea();
END_IF
IF vio_TcpLimitArea.bActive THEN
	vio_Visu.m_SetTcpLimitArea(vi_lr_XMin := vio_TcpLimitArea.fXMin, vi_lr_XMax := vio_TcpLimitArea.fXMax,
		vi_lr_YMin := vio_TcpLimitArea.fYMin, vi_lr_YMax := vio_TcpLimitArea.fYMax,
		vi_lr_ZMin := vio_TcpLimitArea.fZMin, vi_lr_ZMax := vio_TcpLimitArea.fZMax);
ELSE
	vio_Visu.m_ClearTcpLimitArea();
END_IF
END_METHOD

(****************************************************************************************************<br>
© Syntegon Group.<br>
All rights reserved, also regarding any disposal, exploitation, reproduction, editing, distribution,<br>
as well as in the event of applications for industrial property rights.<br>
*****************************************************************************************************<br>
DESCRIPTION:<br>
Passes the effective track modules on to an XTS track's Syn_Visu FB (XTS gantry, XTS loop). Syn_Visu's module<br>
count only grows: the modules are cleared first only when the set has fewer than the visualisation, so its<br>
config version only changes when a value does.<br>
****************************************************************************************************)
METHOD PROTECTED m_PassOnModules : BOOL
VAR_IN_OUT
	vio_Visu							: SynVisu._FB_VisuXtsTrack;	// the track's Syn_Visu FB
END_VAR
VAR_IN_OUT CONSTANT
	(* effective modules *)
	vio_aModules						: ARRAY[0..SynVisu.VISU_GlobalConst_Param.VISU_un_MAX_MODULES - 1] OF SynVisu.ST_VisuTrackModule;
END_VAR
VAR_INPUT
	vi_un_Count							: UINT;	// [-] effective modules in vio_aModules
	vi_un_VisuCount						: UINT;	// [-] modules the visualisation has now, its stConfig.nModuleCount
END_VAR
VAR
	un_TempIndex						: UINT;
END_VAR
m_PassOnModules := TRUE;
IF vi_un_VisuCount > vi_un_Count THEN
	vio_Visu.m_ClearModules();
END_IF
un_TempIndex := 0;
WHILE un_TempIndex < vi_un_Count AND un_TempIndex < SynVisu.VISU_GlobalConst_Param.VISU_un_MAX_MODULES DO
	vio_Visu.m_SetModule(vi_un_Module := un_TempIndex + 1, vi_e_Kind := vio_aModules[un_TempIndex].eKind,
		vi_lr_Length := vio_aModules[un_TempIndex].fLength);
	un_TempIndex := un_TempIndex + 1;
END_WHILE
END_METHOD

(****************************************************************************************************<br>
© Syntegon Group.<br>
All rights reserved, also regarding any disposal, exploitation, reproduction, editing, distribution,<br>
as well as in the event of applications for industrial property rights.<br>
*****************************************************************************************************<br>
DESCRIPTION:<br>
Passes the effective zones on to a Syn_Visu component with zones (robot, detector, station). Syn_Visu's zone<br>
count only grows: the zones are cleared first only when the set has fewer than the visualisation, so its<br>
config version only changes when a value does.<br>
****************************************************************************************************)
METHOD PROTECTED m_PassOnZones : BOOL
VAR_IN_OUT
	vio_Visu							: SynVisu._FB_VisuZoneComponent;	// the component's Syn_Visu FB
END_VAR
VAR_IN_OUT CONSTANT
	(* effective zones *)
	vio_aZones							: ARRAY[0..SynVisu.VISU_GlobalConst_Param.VISU_un_MAX_ZONES - 1] OF SynVisu.ST_VisuZone;
END_VAR
VAR_INPUT
	vi_un_Count							: UINT;	// [-] effective zones in vio_aZones
	vi_un_VisuCount						: UINT;	// [-] zones the visualisation has now, its stConfig.nZoneCount
END_VAR
VAR
	un_TempIndex						: UINT;
END_VAR
m_PassOnZones := TRUE;
IF vi_un_VisuCount > vi_un_Count THEN
	vio_Visu.m_ClearZones();
END_IF
un_TempIndex := 0;
WHILE un_TempIndex < vi_un_Count AND un_TempIndex < SynVisu.VISU_GlobalConst_Param.VISU_un_MAX_ZONES DO
	vio_Visu.m_SetZone(vi_un_Zone := un_TempIndex + 1, vi_udn_ConveyorId := vio_aZones[un_TempIndex].nConveyorId,
		vi_lr_Start := vio_aZones[un_TempIndex].fStart, vi_lr_End := vio_aZones[un_TempIndex].fEnd,
		vi_lr_AllocationOffset := vio_aZones[un_TempIndex].fAllocationOffset,
		vi_lr_CcsOffset := vio_aZones[un_TempIndex].fCcsOffset,
		vi_lr_StartY := vio_aZones[un_TempIndex].fStartY, vi_lr_EndY := vio_aZones[un_TempIndex].fEndY);
	un_TempIndex := un_TempIndex + 1;
END_WHILE
END_METHOD

(****************************************************************************************************<br>
© Syntegon Group.<br>
All rights reserved, also regarding any disposal, exploitation, reproduction, editing, distribution,<br>
as well as in the event of applications for industrial property rights.<br>
*****************************************************************************************************<br>
DESCRIPTION:<br>
Adds this parameter FB to the config manifest under the id of the Syn_Visu component it parametrises.<br>
Idempotent: call it every cycle. The symbol path the gateway reads comes from the instance's own path, as in<br>
Syn_Visu (VISU_un_INSTANCE_PATH_SKIP).<br>
*****************************************************************************************************<br>
OUTPUT VALUES:<br>
FALSE for vi_udn_Id = 0 (but for _FB_ConfigMachine, which registers with id 0), an id already used by a<br>
different entry, or a full manifest.<br>
****************************************************************************************************)
METHOD m_Register : BOOL
VAR_IN_OUT
	vio_Manifest						: ST_ConfigManifest;	// GVL_Config.stManifest of the application
END_VAR
VAR_INPUT
	vi_udn_Id							: UDINT;	// [-] id of the Syn_Visu component, e.g. fb_Infeed.m_Id()
END_VAR
VAR
	e_TempType							: SynVisu.E_VisuComponentType;
	un_TempIndex						: UINT;
END_VAR
m_Register := FALSE;
(* Always report the contract version of the library actually running, also after an online change. *)
vio_Manifest.nProtocolVersion := CONFIG_GlobalConst.CONFIG_un_PROTOCOL_VERSION;
vio_Manifest.sLibraryVersion := CONFIG_GlobalConst.CONFIG_str_LIBRARY_VERSION;
e_TempType := m_ComponentType();
(* Id 0 is the machine FB's, whose type is NONE (_FB_ConfigMachine); every parameter FB has a component's id. *)
IF (vi_udn_Id = 0) <> (e_TempType = SynVisu.E_VisuComponentType.NONE) THEN
	RETURN;
END_IF
IF str_SymbolPath = '' THEN
	str_SymbolPath := m_SymbolPath();
END_IF

(* An existing entry with the same id must match exactly. *)
un_TempIndex := 0;
WHILE un_TempIndex < vio_Manifest.nCount AND un_TempIndex < CONFIG_GlobalConst_Param.CONFIG_un_MAX_MANIFEST_ENTRIES DO
	IF vio_Manifest.aEntries[un_TempIndex].nId = vi_udn_Id THEN
		m_Register := vio_Manifest.aEntries[un_TempIndex].eType = e_TempType
					AND vio_Manifest.aEntries[un_TempIndex].sPath = str_SymbolPath;
		IF m_Register THEN
			udn_ComponentId := vi_udn_Id;
		END_IF
		RETURN;
	END_IF
	un_TempIndex := un_TempIndex + 1;
END_WHILE

(* New entry. *)
IF vio_Manifest.nCount >= CONFIG_GlobalConst_Param.CONFIG_un_MAX_MANIFEST_ENTRIES THEN
	RETURN;
END_IF
vio_Manifest.aEntries[vio_Manifest.nCount].nId := vi_udn_Id;
vio_Manifest.aEntries[vio_Manifest.nCount].eType := e_TempType;
vio_Manifest.aEntries[vio_Manifest.nCount].sPath := str_SymbolPath;
vio_Manifest.nCount := vio_Manifest.nCount + 1;
udn_ComponentId := vi_udn_Id;
m_Register := TRUE;
END_METHOD

(****************************************************************************************************<br>
© Syntegon Group.<br>
All rights reserved, also regarding any disposal, exploitation, reproduction, editing, distribution,<br>
as well as in the event of applications for industrial property rights.<br>
*****************************************************************************************************<br>
DESCRIPTION:<br>
What to do with the staging this cycle: a reset at once; a staged set only while the application allows it<br>
(else the status says PENDING) and only on the active version it is based on (else it is rejected here).<br>
****************************************************************************************************)
METHOD PROTECTED m_Staging : E_ConfigAction
VAR_IN_OUT
	vio_Staging							: ST_ConfigStaging;	// vo_Config.stStaging
	vio_Status							: ST_ConfigStatus;	// vo_Config.stStatus
END_VAR
VAR_INPUT
	vi_b_ApplyAllowed					: BOOL;	// [-] the application allows taking a set over now
	vi_udn_ActiveVersion				: UDINT;	// [-] version of the active set, 0 = program values
END_VAR
m_Staging := E_ConfigAction.NONE;
IF vio_Staging.bReset THEN
	m_Staging := E_ConfigAction.RESET;
ELSIF vio_Staging.bStaged THEN
	IF NOT vi_b_ApplyAllowed THEN
		vio_Status.eResult := E_ConfigResult.PENDING;
	ELSIF vio_Staging.nBaseVersion <> vi_udn_ActiveVersion THEN
		m_Handled(vio_Staging := vio_Staging, vio_Status := vio_Status,
			vi_str_Rejection := CONCAT(CONCAT('Based on version ', UDINT_TO_STRING(vio_Staging.nBaseVersion)),
				CONCAT(', but version ', CONCAT(UDINT_TO_STRING(vi_udn_ActiveVersion), ' is active'))));
	ELSE
		m_Staging := E_ConfigAction.TAKE_OVER;
	END_IF
END_IF
END_METHOD

(****************************************************************************************************<br>
© Syntegon Group.<br>
All rights reserved, also regarding any disposal, exploitation, reproduction, editing, distribution,<br>
as well as in the event of applications for industrial property rights.<br>
*****************************************************************************************************<br>
DESCRIPTION:<br>
Symbol path of this instance's vo_Config as the gateway reads it, from the instance path TwinCAT sets: the<br>
first VISU_un_INSTANCE_PATH_SKIP segments (TwinCAT project, PLC project) are left out, '.vo_Config' is appended.<br>
E.g. 'RPP_Visu.Syn_Visu_Demo.P_VisuDemoDelta.fb_InfeedParam' -> 'P_VisuDemoDelta.fb_InfeedParam.vo_Config'.<br>
****************************************************************************************************)
METHOD PRIVATE m_SymbolPath : STRING(255)
VAR
	un_TempRead							: UINT;	// [-] byte index in str_InstancePath
	un_TempWrite						: UINT;	// [-] byte index in the result
	un_TempDots							: UINT;	// [-] dots passed
END_VAR
VAR CONSTANT
	un_MAX_INDEX						: UINT := 255;	// [-] last byte of a STRING(255), its terminating zero
	by_DOT								: BYTE := 16#2E;	// '.'
	str_SUFFIX							: STRING(15) := '.vo_Config';	// every parameter FB's contract structure
END_VAR
(* Skip the leading segments, up to and including the VISU_un_INSTANCE_PATH_SKIP-th dot. *)
un_TempRead := 0;
un_TempDots := 0;
WHILE un_TempDots < SynVisu.VISU_GlobalConst_Param.VISU_un_INSTANCE_PATH_SKIP AND un_TempRead < un_MAX_INDEX
	AND str_InstancePath[un_TempRead] <> 0
DO
	IF str_InstancePath[un_TempRead] = by_DOT THEN
		un_TempDots := un_TempDots + 1;
	END_IF
	un_TempRead := un_TempRead + 1;
END_WHILE
IF un_TempDots < SynVisu.VISU_GlobalConst_Param.VISU_un_INSTANCE_PATH_SKIP THEN
	un_TempRead := 0;
END_IF

(* The rest of the instance path, then the contract structure. *)
un_TempWrite := 0;
WHILE un_TempRead < un_MAX_INDEX AND str_InstancePath[un_TempRead] <> 0 AND un_TempWrite < un_MAX_INDEX DO
	m_SymbolPath[un_TempWrite] := str_InstancePath[un_TempRead];
	un_TempRead := un_TempRead + 1;
	un_TempWrite := un_TempWrite + 1;
END_WHILE
un_TempRead := 0;
WHILE str_SUFFIX[un_TempRead] <> 0 AND un_TempWrite < un_MAX_INDEX DO
	m_SymbolPath[un_TempWrite] := str_SUFFIX[un_TempRead];
	un_TempRead := un_TempRead + 1;
	un_TempWrite := un_TempWrite + 1;
END_WHILE
m_SymbolPath[un_TempWrite] := 0;
END_METHOD

END_FUNCTION_BLOCK

// POUs/_FB_ConfigConveyor
(****************************************************************************************************<br>
© Syntegon Group.<br>
All rights reserved, also regarding any disposal, exploitation, reproduction, editing, distribution,<br>
as well as in the event of applications for industrial property rights.<br>
*****************************************************************************************************<br>
DESCRIPTION:<br>
Parameter set of one conveyor (ADR 0017): its pose, origin shift and product types, written by the configurator,<br>
taken over when the application allows it. Typical cycle, before the Syn_Visu calls of the conveyor:<br>
  fb_InfeedParam.m_Register(vio_Manifest := GVL_Config.stManifest, vi_udn_Id := fb_Infeed.m_Id());<br>
  fb_InfeedParam.m_Cycle(vio_Default := InfeedDefault, vio_Set := InfeedSet, vi_b_ApplyAllowed := b_Stopped);<br>
  fb_Infeed.m_Configure(vi_Pose := fb_InfeedParam.m_Pose(), vi_lr_Length := 3000, vi_lr_Width := 400);<br>
  fb_InfeedParam.m_PassOn(vio_Visu := fb_Infeed);<br>
InfeedSet is the application's VAR PERSISTENT ST_ConfigConveyorSet; InfeedDefault its program values.<br>
*****************************************************************************************************<br>
OUTPUT VALUES:<br>
vo_Config is the contract structure the gateway reads and writes at the path in the config manifest.<br>
*****************************************************************************************************<br>
VERSION         ¦ DATE       ¦ NAME      ¦ CHANGE<br>
Syn_Config 1.0.0 ¦ 2026-11-10 ¦ J.Willner ¦ First version<br>
****************************************************************************************************)
FUNCTION_BLOCK _FB_ConfigConveyor EXTENDS _FB_ConfigComponent
VAR_OUTPUT
	vo_Config							: ST_ConfigConveyor;	// contract structure of the gateway
END_VAR

(****************************************************************************************************<br>
© Syntegon Group.<br>
All rights reserved, also regarding any disposal, exploitation, reproduction, editing, distribution,<br>
as well as in the event of applications for industrial property rights.<br>
*****************************************************************************************************<br>
DESCRIPTION:<br>
All effective values (origin shift, product types, ...), for the application's own logic.<br>
****************************************************************************************************)
METHOD m_Active : ST_ConfigConveyorParam
m_Active := vo_Config.stActive;
END_METHOD

(****************************************************************************************************<br>
© Syntegon Group.<br>
All rights reserved, also regarding any disposal, exploitation, reproduction, editing, distribution,<br>
as well as in the event of applications for industrial property rights.<br>
*****************************************************************************************************<br>
DESCRIPTION:<br>
A conveyor.<br>
****************************************************************************************************)
METHOD PROTECTED m_ComponentType : SynVisu.E_VisuComponentType
m_ComponentType := SynVisu.E_VisuComponentType.CONVEYOR;
END_METHOD

(****************************************************************************************************<br>
© Syntegon Group.<br>
All rights reserved, also regarding any disposal, exploitation, reproduction, editing, distribution,<br>
as well as in the event of applications for industrial property rights.<br>
*****************************************************************************************************<br>
DESCRIPTION:<br>
Every cycle: handles a staged set or a reset (a set only while vi_b_ApplyAllowed), keeps the active set in<br>
vio_Set and gives the effective values in vo_Config.stActive: the active set while one is valid, else the<br>
program values vio_Default.<br>
*****************************************************************************************************<br>
OUTPUT VALUES:<br>
TRUE in the cycle a set was taken over or reset.<br>
****************************************************************************************************)
METHOD m_Cycle : BOOL
VAR_IN_OUT CONSTANT
	vio_Default							: ST_ConfigConveyorParam;	// the application's program values
END_VAR
VAR_IN_OUT
	vio_Set								: ST_ConfigConveyorSet;	// the application's VAR PERSISTENT active set
END_VAR
VAR_INPUT
	vi_b_ApplyAllowed					: BOOL;	// [-] a staged set may be taken over now, e.g. while the machine stands
END_VAR
VAR
	str_TempRejection					: STRING(80);
END_VAR
m_Cycle := FALSE;
CASE m_Staging(vio_Staging := vo_Config.stStaging, vio_Status := vo_Config.stStatus, vi_b_ApplyAllowed := vi_b_ApplyAllowed,
	vi_udn_ActiveVersion := SEL(vio_Set.bValid, 0, vio_Set.nVersion)) OF
	E_ConfigAction.RESET:
		vio_Set.bValid := FALSE;
		m_Handled(vio_Staging := vo_Config.stStaging, vio_Status := vo_Config.stStatus, vi_str_Rejection := '');
		m_Cycle := TRUE;
	E_ConfigAction.TAKE_OVER:
		str_TempRejection := m_Invalid(vio_Param := vo_Config.stStaged);
		IF str_TempRejection = '' THEN
			vio_Set.nLastVersion := vio_Set.nLastVersion + 1;
			vio_Set.nVersion := vio_Set.nLastVersion;
			vio_Set.stParam := vo_Config.stStaged;
			vio_Set.bValid := TRUE;
			m_Cycle := TRUE;
		END_IF
		m_Handled(vio_Staging := vo_Config.stStaging, vio_Status := vo_Config.stStatus, vi_str_Rejection := str_TempRejection);
END_CASE


(****************************************************************************************************
EFFECTIVE VALUES
****************************************************************************************************)
IF vio_Set.bValid THEN
	vo_Config.stActive := vio_Set.stParam;
	vo_Config.stStatus.nActiveVersion := vio_Set.nVersion;
ELSE
	vo_Config.stActive := vio_Default;
	vo_Config.stStatus.nActiveVersion := 0;
END_IF
END_METHOD

(****************************************************************************************************<br>
© Syntegon Group.<br>
All rights reserved, also regarding any disposal, exploitation, reproduction, editing, distribution,<br>
as well as in the event of applications for industrial property rights.<br>
*****************************************************************************************************<br>
DESCRIPTION:<br>
Why a staged set cannot be taken over; '' when it can: more product types than the list holds, a product type<br>
without a number or a number used twice.<br>
****************************************************************************************************)
METHOD PRIVATE m_Invalid : STRING(80)
VAR_IN_OUT CONSTANT
	vio_Param							: ST_ConfigConveyorParam;	// the staged set
END_VAR
VAR
	un_TempIndex						: UINT;
	un_TempOther						: UINT;
END_VAR
m_Invalid := '';
IF vio_Param.nProductTypeCount > SynVisu.VISU_GlobalConst_Param.VISU_un_MAX_PRODUCT_TYPES THEN
	m_Invalid := CONCAT('More than ', CONCAT(UINT_TO_STRING(SynVisu.VISU_GlobalConst_Param.VISU_un_MAX_PRODUCT_TYPES), ' product types'));
	RETURN;
END_IF
un_TempIndex := 0;
WHILE un_TempIndex < vio_Param.nProductTypeCount DO
	IF vio_Param.aProductTypes[un_TempIndex].nId = 0 THEN
		m_Invalid := 'A product type without a number';
		RETURN;
	END_IF
	un_TempOther := 0;
	WHILE un_TempOther < un_TempIndex DO
		IF vio_Param.aProductTypes[un_TempOther].nId = vio_Param.aProductTypes[un_TempIndex].nId THEN
			m_Invalid := CONCAT('Product type ', CONCAT(UDINT_TO_STRING(vio_Param.aProductTypes[un_TempIndex].nId), ' is defined twice'));
			RETURN;
		END_IF
		un_TempOther := un_TempOther + 1;
	END_WHILE
	un_TempIndex := un_TempIndex + 1;
END_WHILE
END_METHOD

(****************************************************************************************************<br>
© Syntegon Group.<br>
All rights reserved, also regarding any disposal, exploitation, reproduction, editing, distribution,<br>
as well as in the event of applications for industrial property rights.<br>
*****************************************************************************************************<br>
DESCRIPTION:<br>
Passes the effective origin shift and product types on to the conveyor's Syn_Visu FB, so the visualisation shows<br>
what the machine uses. The pose goes with the application's own m_Configure call (with the belt's length and<br>
width, hardware): vi_Pose := m_Pose(). Call it after m_Cycle, every cycle; Syn_Visu's config version only<br>
changes when a value does.<br>
*****************************************************************************************************<br>
LIMITS:<br>
Syn_Visu cannot remove a product type: one the set no longer has stays in the visualisation until the<br>
application restarts (the configurator warns of the difference).<br>
****************************************************************************************************)
METHOD m_PassOn : BOOL
VAR_IN_OUT
	vio_Visu							: SynVisu._FB_VisuConveyor;	// the conveyor's Syn_Visu FB
END_VAR
VAR
	un_TempIndex						: UINT;
END_VAR
m_PassOn := TRUE;
vio_Visu.m_SetOriginShift(vi_lr_X := vo_Config.stActive.stOriginShift.fX, vi_lr_Y := vo_Config.stActive.stOriginShift.fY,
	vi_lr_Z := vo_Config.stActive.stOriginShift.fZ);
un_TempIndex := 0;
WHILE un_TempIndex < vo_Config.stActive.nProductTypeCount
	AND un_TempIndex < SynVisu.VISU_GlobalConst_Param.VISU_un_MAX_PRODUCT_TYPES
DO
	vio_Visu.m_SetProductType(vi_udn_Id := vo_Config.stActive.aProductTypes[un_TempIndex].nId,
		vi_lr_Length := vo_Config.stActive.aProductTypes[un_TempIndex].fLength,
		vi_lr_Width := vo_Config.stActive.aProductTypes[un_TempIndex].fWidth,
		vi_lr_Height := vo_Config.stActive.aProductTypes[un_TempIndex].fHeight,
		vi_e_Shape := vo_Config.stActive.aProductTypes[un_TempIndex].eShape,
		vi_lr_CornerRadius := vo_Config.stActive.aProductTypes[un_TempIndex].fCornerRadius);
	un_TempIndex := un_TempIndex + 1;
END_WHILE
END_METHOD

(****************************************************************************************************<br>
© Syntegon Group.<br>
All rights reserved, also regarding any disposal, exploitation, reproduction, editing, distribution,<br>
as well as in the event of applications for industrial property rights.<br>
*****************************************************************************************************<br>
DESCRIPTION:<br>
Effective pose of the belt start (MCS), for the application's logic and its Syn_Visu m_Configure call.<br>
****************************************************************************************************)
METHOD m_Pose : SynVisu.ST_VisuPose
m_Pose := vo_Config.stActive.stPose;
END_METHOD

END_FUNCTION_BLOCK

// POUs/_FB_ConfigDelta
(****************************************************************************************************<br>
© Syntegon Group.<br>
All rights reserved, also regarding any disposal, exploitation, reproduction, editing, distribution,<br>
as well as in the event of applications for industrial property rights.<br>
*****************************************************************************************************<br>
DESCRIPTION:<br>
Parameter set of one Delta robot (ADR 0017): its pose, origin shift, zones, gripper fingers, working area,<br>
limit area and TCP limit area, written by the configurator, taken over when the application allows it.<br>
Typical cycle:<br>
  fb_Delta1Param.m_Register(vio_Manifest := GVL_Config.stManifest, vi_udn_Id := fb_Delta1.m_Id());<br>
  fb_Delta1Param.m_Cycle(vio_Default := Delta1Default, vio_Set := Delta1Set, vi_b_ApplyAllowed := b_Stopped);<br>
  fb_Delta1.m_Configure(vi_Pose := fb_Delta1Param.m_Pose(), vi_lr_BaseRadius := 200, ...);<br>
  fb_Delta1Param.m_PassOn(vio_Visu := fb_Delta1);<br>
The application's pick logic takes its zones from m_Zone / m_Active, not from its own constants.<br>
*****************************************************************************************************<br>
OUTPUT VALUES:<br>
vo_Config is the contract structure the gateway reads and writes at the path in the config manifest.<br>
*****************************************************************************************************<br>
VERSION         ¦ DATE       ¦ NAME      ¦ CHANGE<br>
Syn_Config 1.0.0 ¦ 2026-11-10 ¦ J.Willner ¦ First version<br>
Syn_Config 1.1.0 ¦ 2026-11-10 ¦ J.Willner ¦ m_PassOn, m_Invalid through the shared helpers<br>
Syn_Config 2.0.0 ¦ 2026-11-11 ¦ J.Willner ¦ Gripper fingers with their offsets (ADR 0018)<br>
****************************************************************************************************)
FUNCTION_BLOCK _FB_ConfigDelta EXTENDS _FB_ConfigComponent
VAR_OUTPUT
	vo_Config							: ST_ConfigDelta;	// contract structure of the gateway
END_VAR

(****************************************************************************************************<br>
© Syntegon Group.<br>
All rights reserved, also regarding any disposal, exploitation, reproduction, editing, distribution,<br>
as well as in the event of applications for industrial property rights.<br>
*****************************************************************************************************<br>
DESCRIPTION:<br>
All effective values (zones, working and limit areas, ...), for the application's own logic.<br>
****************************************************************************************************)
METHOD m_Active : ST_ConfigDeltaParam
m_Active := vo_Config.stActive;
END_METHOD

(****************************************************************************************************<br>
© Syntegon Group.<br>
All rights reserved, also regarding any disposal, exploitation, reproduction, editing, distribution,<br>
as well as in the event of applications for industrial property rights.<br>
*****************************************************************************************************<br>
DESCRIPTION:<br>
A Delta robot.<br>
****************************************************************************************************)
METHOD PROTECTED m_ComponentType : SynVisu.E_VisuComponentType
m_ComponentType := SynVisu.E_VisuComponentType.DELTA;
END_METHOD

(****************************************************************************************************<br>
© Syntegon Group.<br>
All rights reserved, also regarding any disposal, exploitation, reproduction, editing, distribution,<br>
as well as in the event of applications for industrial property rights.<br>
*****************************************************************************************************<br>
DESCRIPTION:<br>
Every cycle: handles a staged set or a reset (a set only while vi_b_ApplyAllowed), keeps the active set in<br>
vio_Set and gives the effective values in vo_Config.stActive: the active set while one is valid, else the<br>
program values vio_Default.<br>
*****************************************************************************************************<br>
OUTPUT VALUES:<br>
TRUE in the cycle a set was taken over or reset.<br>
****************************************************************************************************)
METHOD m_Cycle : BOOL
VAR_IN_OUT CONSTANT
	vio_Default							: ST_ConfigDeltaParam;	// the application's program values
END_VAR
VAR_IN_OUT
	vio_Set								: ST_ConfigDeltaSet;	// the application's VAR PERSISTENT active set
END_VAR
VAR_INPUT
	vi_b_ApplyAllowed					: BOOL;	// [-] a staged set may be taken over now, e.g. while the machine stands
END_VAR
VAR
	str_TempRejection					: STRING(80);
END_VAR
m_Cycle := FALSE;
CASE m_Staging(vio_Staging := vo_Config.stStaging, vio_Status := vo_Config.stStatus, vi_b_ApplyAllowed := vi_b_ApplyAllowed,
	vi_udn_ActiveVersion := SEL(vio_Set.bValid, 0, vio_Set.nVersion)) OF
	E_ConfigAction.RESET:
		vio_Set.bValid := FALSE;
		m_Handled(vio_Staging := vo_Config.stStaging, vio_Status := vo_Config.stStatus, vi_str_Rejection := '');
		m_Cycle := TRUE;
	E_ConfigAction.TAKE_OVER:
		str_TempRejection := m_Invalid(vio_Param := vo_Config.stStaged);
		IF str_TempRejection = '' THEN
			vio_Set.nLastVersion := vio_Set.nLastVersion + 1;
			vio_Set.nVersion := vio_Set.nLastVersion;
			vio_Set.stParam := vo_Config.stStaged;
			vio_Set.bValid := TRUE;
			m_Cycle := TRUE;
		END_IF
		m_Handled(vio_Staging := vo_Config.stStaging, vio_Status := vo_Config.stStatus, vi_str_Rejection := str_TempRejection);
END_CASE


(****************************************************************************************************
EFFECTIVE VALUES
****************************************************************************************************)
IF vio_Set.bValid THEN
	vo_Config.stActive := vio_Set.stParam;
	vo_Config.stStatus.nActiveVersion := vio_Set.nVersion;
ELSE
	vo_Config.stActive := vio_Default;
	vo_Config.stStatus.nActiveVersion := 0;
END_IF
END_METHOD

(****************************************************************************************************<br>
© Syntegon Group.<br>
All rights reserved, also regarding any disposal, exploitation, reproduction, editing, distribution,<br>
as well as in the event of applications for industrial property rights.<br>
*****************************************************************************************************<br>
DESCRIPTION:<br>
Why a staged set cannot be taken over; '' when it can: more zones or fingers than the lists hold, a zone on no<br>
conveyor (id 0), or a finger without a diameter or height.<br>
****************************************************************************************************)
METHOD PRIVATE m_Invalid : STRING(80)
VAR_IN_OUT CONSTANT
	vio_Param							: ST_ConfigDeltaParam;	// the staged set
END_VAR
m_Invalid := m_InvalidZones(vio_aZones := vio_Param.aZones, vi_un_Count := vio_Param.nZoneCount);
IF m_Invalid = '' THEN
	m_Invalid := m_InvalidFingers(vio_aFingers := vio_Param.aFingers, vi_un_Count := vio_Param.nFingerCount);
END_IF
END_METHOD

(****************************************************************************************************<br>
© Syntegon Group.<br>
All rights reserved, also regarding any disposal, exploitation, reproduction, editing, distribution,<br>
as well as in the event of applications for industrial property rights.<br>
*****************************************************************************************************<br>
DESCRIPTION:<br>
Passes the effective origin shift, working area, limit areas, zones and fingers on to the Delta's Syn_Visu<br>
FB, so the visualisation shows what the machine uses. The pose goes with the application's own m_Configure<br>
call (with the arm geometry, hardware): vi_Pose := m_Pose(). Call it after m_Cycle, every cycle; Syn_Visu's<br>
config version only changes when a value does (zones and fingers are cleared only when the set has fewer than<br>
the visualisation).<br>
****************************************************************************************************)
METHOD m_PassOn : BOOL
VAR_IN_OUT
	vio_Visu							: SynVisu._FB_VisuDelta;	// the Delta's Syn_Visu FB
END_VAR
m_PassOn := TRUE;
vio_Visu.m_SetOriginShift(vi_lr_X := vo_Config.stActive.stOriginShift.fX, vi_lr_Y := vo_Config.stActive.stOriginShift.fY,
	vi_lr_Z := vo_Config.stActive.stOriginShift.fZ);
vio_Visu.m_SetWorkingArea(vi_lr_Radius := vo_Config.stActive.stWorkingArea.fRadius,
	vi_lr_ZMin := vo_Config.stActive.stWorkingArea.fZMin, vi_lr_ZMax := vo_Config.stActive.stWorkingArea.fZMax,
	vi_lr_ConeHeight := vo_Config.stActive.stWorkingArea.fConeHeight,
	vi_lr_ConeBottomRadius := vo_Config.stActive.stWorkingArea.fConeBottomRadius);
m_PassOnLimitAreas(vio_Visu := vio_Visu, vio_LimitArea := vo_Config.stActive.stLimitArea,
	vio_TcpLimitArea := vo_Config.stActive.stTcpLimitArea);
m_PassOnZones(vio_Visu := vio_Visu, vio_aZones := vo_Config.stActive.aZones, vi_un_Count := vo_Config.stActive.nZoneCount,
	vi_un_VisuCount := vio_Visu.vo_Visu.stConfig.nZoneCount);
m_PassOnFingers(vio_Visu := vio_Visu, vio_aFingers := vo_Config.stActive.aFingers,
	vi_un_Count := vo_Config.stActive.nFingerCount, vi_un_VisuCount := vio_Visu.vo_Visu.stConfig.nFingerCount);
END_METHOD

(****************************************************************************************************<br>
© Syntegon Group.<br>
All rights reserved, also regarding any disposal, exploitation, reproduction, editing, distribution,<br>
as well as in the event of applications for industrial property rights.<br>
*****************************************************************************************************<br>
DESCRIPTION:<br>
Effective pose of the base centre (MCS), for the application's logic and its Syn_Visu m_Configure call.<br>
****************************************************************************************************)
METHOD m_Pose : SynVisu.ST_VisuPose
m_Pose := vo_Config.stActive.stPose;
END_METHOD

(****************************************************************************************************<br>
© Syntegon Group.<br>
All rights reserved, also regarding any disposal, exploitation, reproduction, editing, distribution,<br>
as well as in the event of applications for industrial property rights.<br>
*****************************************************************************************************<br>
DESCRIPTION:<br>
Effective zone vi_un_Zone (1-based, as in Syn_Visu's m_SetZone), for the application's pick and place logic.<br>
*****************************************************************************************************<br>
OUTPUT VALUES:<br>
A zone with nConveyorId = 0 for a number outside 1..m_ZoneCount().<br>
****************************************************************************************************)
METHOD m_Zone : SynVisu.ST_VisuZone
VAR_INPUT
	vi_un_Zone							: UINT;	// [-] 1-based
END_VAR
IF vi_un_Zone >= 1 AND vi_un_Zone <= vo_Config.stActive.nZoneCount
	AND vi_un_Zone <= SynVisu.VISU_GlobalConst_Param.VISU_un_MAX_ZONES
THEN
	m_Zone := vo_Config.stActive.aZones[vi_un_Zone - 1];
END_IF
END_METHOD

(****************************************************************************************************<br>
© Syntegon Group.<br>
All rights reserved, also regarding any disposal, exploitation, reproduction, editing, distribution,<br>
as well as in the event of applications for industrial property rights.<br>
*****************************************************************************************************<br>
DESCRIPTION:<br>
Number of effective zones.<br>
****************************************************************************************************)
METHOD m_ZoneCount : UINT
m_ZoneCount := vo_Config.stActive.nZoneCount;
END_METHOD

END_FUNCTION_BLOCK

// POUs/_FB_ConfigXtsGantry
(****************************************************************************************************<br>
© Syntegon Group.<br>
All rights reserved, also regarding any disposal, exploitation, reproduction, editing, distribution,<br>
as well as in the event of applications for industrial property rights.<br>
*****************************************************************************************************<br>
DESCRIPTION:<br>
Parameter set of one XTS gantry (ADR 0017): its pose, origin shift, track modules, zones, gripper fingers,<br>
limit area and TCP limit area, written by the configurator, taken over when the application allows it.<br>
Typical cycle:<br>
  fb_IdhParam.m_Register(vio_Manifest := GVL_Config.stManifest, vi_udn_Id := fb_Idh.m_Id());<br>
  fb_IdhParam.m_Cycle(vio_Default := IdhDefault, vio_Set := IdhSet, vi_b_ApplyAllowed := b_Stopped);<br>
  fb_Idh.m_Configure(vi_Pose := fb_IdhParam.m_Pose(), vi_lr_XMin := 0, ...);<br>
  fb_IdhParam.m_PassOn(vio_Visu := fb_Idh);<br>
The application's logic takes its track and zones from m_Active, not from its own constants.<br>
*****************************************************************************************************<br>
OUTPUT VALUES:<br>
vo_Config is the contract structure the gateway reads and writes at the path in the config manifest.<br>
*****************************************************************************************************<br>
VERSION         ¦ DATE       ¦ NAME      ¦ CHANGE<br>
Syn_Config 1.1.0 ¦ 2026-11-10 ¦ J.Willner ¦ New<br>
Syn_Config 2.0.0 ¦ 2026-11-11 ¦ J.Willner ¦ Gripper fingers with their offsets (ADR 0018)<br>
****************************************************************************************************)
FUNCTION_BLOCK _FB_ConfigXtsGantry EXTENDS _FB_ConfigComponent
VAR_OUTPUT
	vo_Config							: ST_ConfigXtsGantry;	// contract structure of the gateway
END_VAR

(****************************************************************************************************<br>
© Syntegon Group.<br>
All rights reserved, also regarding any disposal, exploitation, reproduction, editing, distribution,<br>
as well as in the event of applications for industrial property rights.<br>
*****************************************************************************************************<br>
DESCRIPTION:<br>
All effective values (track modules, zones, limit areas, ...), for the application's own logic.<br>
****************************************************************************************************)
METHOD m_Active : ST_ConfigXtsGantryParam
m_Active := vo_Config.stActive;
END_METHOD

(****************************************************************************************************<br>
© Syntegon Group.<br>
All rights reserved, also regarding any disposal, exploitation, reproduction, editing, distribution,<br>
as well as in the event of applications for industrial property rights.<br>
*****************************************************************************************************<br>
DESCRIPTION:<br>
An XTS gantry.<br>
****************************************************************************************************)
METHOD PROTECTED m_ComponentType : SynVisu.E_VisuComponentType
m_ComponentType := SynVisu.E_VisuComponentType.XTS_GANTRY;
END_METHOD

(****************************************************************************************************<br>
© Syntegon Group.<br>
All rights reserved, also regarding any disposal, exploitation, reproduction, editing, distribution,<br>
as well as in the event of applications for industrial property rights.<br>
*****************************************************************************************************<br>
DESCRIPTION:<br>
Every cycle: handles a staged set or a reset (a set only while vi_b_ApplyAllowed), keeps the active set in<br>
vio_Set and gives the effective values in vo_Config.stActive: the active set while one is valid, else the<br>
program values vio_Default.<br>
*****************************************************************************************************<br>
OUTPUT VALUES:<br>
TRUE in the cycle a set was taken over or reset.<br>
****************************************************************************************************)
METHOD m_Cycle : BOOL
VAR_IN_OUT CONSTANT
	vio_Default							: ST_ConfigXtsGantryParam;	// the application's program values
END_VAR
VAR_IN_OUT
	vio_Set								: ST_ConfigXtsGantrySet;	// the application's VAR PERSISTENT active set
END_VAR
VAR_INPUT
	vi_b_ApplyAllowed					: BOOL;	// [-] a staged set may be taken over now, e.g. while the machine stands
END_VAR
VAR
	str_TempRejection					: STRING(80);
END_VAR
m_Cycle := FALSE;
CASE m_Staging(vio_Staging := vo_Config.stStaging, vio_Status := vo_Config.stStatus, vi_b_ApplyAllowed := vi_b_ApplyAllowed,
	vi_udn_ActiveVersion := SEL(vio_Set.bValid, 0, vio_Set.nVersion)) OF
	E_ConfigAction.RESET:
		vio_Set.bValid := FALSE;
		m_Handled(vio_Staging := vo_Config.stStaging, vio_Status := vo_Config.stStatus, vi_str_Rejection := '');
		m_Cycle := TRUE;
	E_ConfigAction.TAKE_OVER:
		str_TempRejection := m_Invalid(vio_Param := vo_Config.stStaged);
		IF str_TempRejection = '' THEN
			vio_Set.nLastVersion := vio_Set.nLastVersion + 1;
			vio_Set.nVersion := vio_Set.nLastVersion;
			vio_Set.stParam := vo_Config.stStaged;
			vio_Set.bValid := TRUE;
			m_Cycle := TRUE;
		END_IF
		m_Handled(vio_Staging := vo_Config.stStaging, vio_Status := vo_Config.stStatus, vi_str_Rejection := str_TempRejection);
END_CASE


(****************************************************************************************************
EFFECTIVE VALUES
****************************************************************************************************)
IF vio_Set.bValid THEN
	vo_Config.stActive := vio_Set.stParam;
	vo_Config.stStatus.nActiveVersion := vio_Set.nVersion;
ELSE
	vo_Config.stActive := vio_Default;
	vo_Config.stStatus.nActiveVersion := 0;
END_IF
END_METHOD

(****************************************************************************************************<br>
© Syntegon Group.<br>
All rights reserved, also regarding any disposal, exploitation, reproduction, editing, distribution,<br>
as well as in the event of applications for industrial property rights.<br>
*****************************************************************************************************<br>
DESCRIPTION:<br>
Why a staged set cannot be taken over; '' when it can: a track without modules, more modules, zones or fingers<br>
than the lists hold, a module without a length, a zone on no conveyor (id 0), or a finger without a diameter or<br>
height.<br>
****************************************************************************************************)
METHOD PRIVATE m_Invalid : STRING(80)
VAR_IN_OUT CONSTANT
	vio_Param							: ST_ConfigXtsGantryParam;	// the staged set
END_VAR
m_Invalid := m_InvalidModules(vio_aModules := vio_Param.aModules, vi_un_Count := vio_Param.nModuleCount);
IF m_Invalid = '' THEN
	m_Invalid := m_InvalidZones(vio_aZones := vio_Param.aZones, vi_un_Count := vio_Param.nZoneCount);
END_IF
IF m_Invalid = '' THEN
	m_Invalid := m_InvalidFingers(vio_aFingers := vio_Param.aFingers, vi_un_Count := vio_Param.nFingerCount);
END_IF
END_METHOD

(****************************************************************************************************<br>
© Syntegon Group.<br>
All rights reserved, also regarding any disposal, exploitation, reproduction, editing, distribution,<br>
as well as in the event of applications for industrial property rights.<br>
*****************************************************************************************************<br>
DESCRIPTION:<br>
Passes the effective origin shift, track modules, limit areas, zones and fingers on to the gantry's Syn_Visu<br>
FB, so the visualisation shows what the machine uses. The pose goes with the application's own m_Configure<br>
call (with the strokes and tool offsets, hardware): vi_Pose := m_Pose(). Call it after m_Cycle, every cycle;<br>
Syn_Visu's config version only changes when a value does.<br>
****************************************************************************************************)
METHOD m_PassOn : BOOL
VAR_IN_OUT
	vio_Visu							: SynVisu._FB_VisuXtsGantry;	// the gantry's Syn_Visu FB
END_VAR
m_PassOn := TRUE;
vio_Visu.m_SetOriginShift(vi_lr_X := vo_Config.stActive.stOriginShift.fX, vi_lr_Y := vo_Config.stActive.stOriginShift.fY,
	vi_lr_Z := vo_Config.stActive.stOriginShift.fZ);
m_PassOnModules(vio_Visu := vio_Visu, vio_aModules := vo_Config.stActive.aModules,
	vi_un_Count := vo_Config.stActive.nModuleCount, vi_un_VisuCount := vio_Visu.vo_Visu.stConfig.nModuleCount);
m_PassOnLimitAreas(vio_Visu := vio_Visu, vio_LimitArea := vo_Config.stActive.stLimitArea,
	vio_TcpLimitArea := vo_Config.stActive.stTcpLimitArea);
m_PassOnZones(vio_Visu := vio_Visu, vio_aZones := vo_Config.stActive.aZones, vi_un_Count := vo_Config.stActive.nZoneCount,
	vi_un_VisuCount := vio_Visu.vo_Visu.stConfig.nZoneCount);
m_PassOnFingers(vio_Visu := vio_Visu, vio_aFingers := vo_Config.stActive.aFingers,
	vi_un_Count := vo_Config.stActive.nFingerCount, vi_un_VisuCount := vio_Visu.vo_Visu.stConfig.nFingerCount);
END_METHOD

(****************************************************************************************************<br>
© Syntegon Group.<br>
All rights reserved, also regarding any disposal, exploitation, reproduction, editing, distribution,<br>
as well as in the event of applications for industrial property rights.<br>
*****************************************************************************************************<br>
DESCRIPTION:<br>
Effective pose of the track start (MCS), for the application's logic and its Syn_Visu m_Configure call.<br>
****************************************************************************************************)
METHOD m_Pose : SynVisu.ST_VisuPose
m_Pose := vo_Config.stActive.stPose;
END_METHOD

END_FUNCTION_BLOCK

// POUs/_FB_ConfigMachine
(****************************************************************************************************<br>
© Syntegon Group.<br>
All rights reserved, also regarding any disposal, exploitation, reproduction, editing, distribution,<br>
as well as in the event of applications for industrial property rights.<br>
*****************************************************************************************************<br>
DESCRIPTION:<br>
The machine as a whole (config protocol 3, ADR 0022): the recipe fields the application declares (process values<br>
such as belt speed, picks per cycle, the product pattern), their staging by the Simulator with the mechanism of the<br>
parameter sets, and the machine commands Start, Stop and Reset the application answers. One per application,<br>
listed in the config manifest with id 0. Typical cycle:<br>
  fb_Machine.m_Register(vio_Manifest := GVL_Config.stManifest, vi_udn_Id := 0);<br>
  fb_Machine.m_DeclareField(vi_un_Field := 1, vi_str_Name := 'BeltSpeed', vi_udn_Group := fb_Infeed.m_Id(),<br>
    vi_e_Type := E_ConfigFieldType.NUMBER, vi_str_Unit := 'mm/s', vi_lr_Min := 0, vi_lr_Max := 500,<br>
    vi_lr_ProgramValue := 150);<br>
  fb_Machine.m_Cycle(vio_Set := RecipeSet, vi_b_ApplyAllowed := b_Stopped);<br>
  lr_BeltSpeed := fb_Machine.m_Value(vi_un_Field := 1);<br>
  CASE fb_Machine.m_Command() OF E_ConfigCommand.START: ...<br>
    fb_Machine.m_AnswerCommand(vi_b_Accepted := TRUE, vi_str_Reason := ''); END_CASE<br>
RecipeSet is the application's VAR PERSISTENT ST_ConfigRecipeSet.<br>
*****************************************************************************************************<br>
OUTPUT VALUES:<br>
vo_Config is the contract structure the gateway reads and writes at the path in the config manifest.<br>
*****************************************************************************************************<br>
LIMITS:<br>
CONFIG_un_MAX_RECIPE_FIELDS fields, CONFIG_un_MAX_CHOICES choices each. The gateway reads the declarations when<br>
it discovers the PLC: declare every field from the start and keep their order.<br>
*****************************************************************************************************<br>
VERSION         ¦ DATE       ¦ NAME      ¦ CHANGE<br>
Syn_Config 2.1.0 ¦ 2026-11-14 ¦ J.Willner ¦ Created: recipe fields and machine commands (protocol 3)<br>
****************************************************************************************************)
FUNCTION_BLOCK _FB_ConfigMachine EXTENDS _FB_ConfigComponent
VAR_OUTPUT
	vo_Config							: ST_ConfigMachine;	// contract structure of the gateway
END_VAR

(****************************************************************************************************<br>
© Syntegon Group.<br>
All rights reserved, also regarding any disposal, exploitation, reproduction, editing, distribution,<br>
as well as in the event of applications for industrial property rights.<br>
*****************************************************************************************************<br>
DESCRIPTION:<br>
Answers the waiting machine command: accepted, or rejected with the reason the Simulator shows. The command no<br>
longer waits afterwards.<br>
*****************************************************************************************************<br>
OUTPUT VALUES:<br>
FALSE while no command waits.<br>
****************************************************************************************************)
METHOD m_AnswerCommand : BOOL
VAR_INPUT
	vi_b_Accepted						: BOOL;	// TRUE: the application carries the command out
	vi_str_Reason						: STRING(80);	// why it is rejected, '' when accepted
END_VAR
m_AnswerCommand := vo_Config.stCommand.bRequested;
IF NOT m_AnswerCommand THEN
	RETURN;
END_IF
vo_Config.stCommandStatus.nHandledCommandId := vo_Config.stCommand.nCommandId;
vo_Config.stCommandStatus.eResult := SEL(vi_b_Accepted, E_ConfigCommandResult.REJECTED, E_ConfigCommandResult.ACCEPTED);
vo_Config.stCommandStatus.sMessage := SEL(vi_b_Accepted, vi_str_Reason, '');
vo_Config.stCommand.bRequested := FALSE;
END_METHOD

